(* IEC 61131-3 sources: daoli-st-library/DL_Motion (part 7) *)

(* ---- FB_DL_AxisInertiaIdent.st ---- *)
(*==============================================================================
 * 组件名称 (Component)  : FB_DL_AxisInertiaIdent
 * 所属子库 (Sublibrary) : DL_Motion
 * 当前版本 (Version)    : 1.0.0
 * 兼容性   (Platform)   : CODESYS 3.5+ / TwinCAT 3 / 汇川 InoProShop / 施耐德 Machine Expert
 *                         仅依赖 Standard.library（R_TRIG / ABS）与库内开方内核 FC_DL_SqrtEx，
 *                         零厂商私有库
 * 功能描述 (Function)   : 转动惯量与摩擦转矩在线辨识。在加速段采集 (a, T) 样本对，用最小二乘
 *                         闭式解拟合 T = J·a + Tf，得惯量 J 与摩擦转矩 Tf：
 *                         J = 〔n·ΣaT − Σa·ΣT〕/〔n·Σa² − (Σa)²〕，Tf = 〔ΣT − J·Σa〕/ n。
 *                         采样门限：|fAcc| >= fAccMin 才纳入样本；有效样本数 < nSampleMin 不出结果。
 *                         置信度：残差均方根 fRms 超 fRmsMax 时 bConfident = FALSE——**照出结果但标
 *                         不可信**（不静默丢弃，现场需要看到「拟合出来了但不可信」这个事实）。
 *                         bFreeze 为真时停止更新，fInertiaOut 保持（供调试比对）。
 * 接口     (Interface)  : 输入 fAcc 角加速度、fTorque 转矩、fAccMin 采样门限、nSampleMin 最小
 *                         样本数、fRmsMax 残差均方根上限、bEnable 使能、bFreeze 结果冻结、bReset 复位；
 *                         输出 fInertiaOut 惯量、fFrictionOut 摩擦转矩、fRms 残差均方根、
 *                         bConfident 置信标记、nSampleCount 有效样本数、eState / eCause / bError / nErrId。
 * 边界     (Boundary)   : ① 回归分母〔n·Σa² − (Σa)²〕<= DL_FLOAT_EPS 判定样本不可分（如全等
 *                         加速度），置信息级并**保持上次结果**（不清零，避免把「没算出来」错当
 *                         「惯量为 0」）；② 全部累加量用 LREAL 防精度丢失；**本件用累积量闭式解，
 *                         不使用样本环形缓冲**，故无下标越界路径（派单「环缓冲下标先判边界」
 *                         条款以零数组方式结构性满足）；
 *                         ③ 组态闸：fAccMin <= 0.0、nSampleMin = 0、fRmsMax <= 0.0 或任一浮点引脚
 *                         NaN → 故障锁存；④ 输入非有限 → 该样本剔除并计数，不污染累加量；
 *                         ⑤ R_TRIG 一枚段 0 无条件刷新（本件为纯算术拟合，无工艺相计时）；
 *                         ⑥ 故障相迁出唯一路径 = bReset 上升沿；⑦ 零全局耦合（无 GVL / 无物理地址）。
 * 解除式   (Release)    : bReset 上升沿 ∧ 组态合法 ∧ 回归分母非病态（当拍量，R240 范式）。
 *                         自证可满足（终审两式 1）：分母只依赖累加量与样本数，复位后累加量清空
 *                         即重新开始积累，加速度样本一旦分散分母即脱离病态，无恒假因子。
 * 码表     (Codes)      : 16#0004_03B7 故障级：惯量辨识故障总码（组态非法 / 输入非有限累计超限 /
 *                         非法相位），锁存至 bReset 上升沿，归因由 eCause 承载（R190 单件单总码）；
 *                         16#0004_04B7 信息级：非故障台账事件（分母病态保持上次结果 / 样本数不足）。
 *                         加码反证（R90）：二者都不改 bError、不改 eCause，且 bConfident 仍可能为真
 *                         （保持的旧结果可能高置信），若不立码则「本轮没算出新结果」不可观测，故立
 *                         一码；二者共用一码的依据是「都只要求留痕」，区分由 nSampleCount 反推。
 *                         码段说明：0004 段故障子带 03xx / 信息子带 04xx，本件取 03B7 / 04B7
 *                         （源码实扫该两槽为空，续接同子带已用最大值，未回填碎片孔洞）。
 * 开源溯源 (Origin)     : 道莅自研 clean-room（参考最小二乘闭式解与运动辨识参数域，零代码行复制；
 *                         t2-4-s7-motion 族）
 * 修订历史 (Revision)   : 2026-11-19  v1.0.0  R45 首版（批次 3 · 序号 13）
 *==============================================================================*)

TYPE E_DL_AiiState :
(
    eIdle  := 0,     // 失能或样本不足（无结果） / Idle, disabled or not enough samples
    eRun   := 10,    // 辨识运行 / Identification running
    eFault := 90     // 故障锁存相 / Fault latched phase
);
END_TYPE

TYPE E_DL_AiiCause :
(
    eNone       := 0,   // 无故障成因 / No cause
    eCfgIllegal := 1,   // 组态非法 / Illegal configuration
    eNonFinRun  := 2,   // 输入非有限累计超限 / Too many consecutive non-finite inputs
    ePhaseBad   := 3    // 非法相位兜底 / Illegal phase fallback
);
END_TYPE

FUNCTION_BLOCK FB_DL_AxisInertiaIdent
VAR_INPUT
    fAcc        : REAL := 0.0;          // 角加速度（或线加速度） [rad/s²] / Angular acceleration [rad/s2]
    fTorque     : REAL := 0.0;          // 实测转矩 [N·m] / Measured torque [N·m]
    fAccMin     : REAL := 5.0;          // 采样门限（|a| 大于该值才纳入），域 > 0.0 [rad/s²] / Sampling threshold, domain > 0.0 [rad/s2]
    nSampleMin  : UDINT := 50;          // 最小有效样本数，域 > 0 [个] / Minimum sample count, domain > 0 [pcs]
    fRmsMax     : REAL := 0.50;         // 残差均方根上限，域 > 0.0 [N·m] / Residual RMS limit, domain > 0.0 [N·m]
    bEnable     : BOOL := TRUE;         // 辨识使能 [-] / Identification enable
    bFreeze     : BOOL := FALSE;        // 结果冻结（停止更新，保持末值） [-] / Freeze results, hold last value
    bReset      : BOOL := FALSE;        // 复位命令，上升沿清故障并使累加量净重装 [-] / Reset clears fault and re-arms accumulators
END_VAR
VAR_OUTPUT
    fInertiaOut  : REAL;                // 辨识惯量（拟合斜率） [kg·m²] / Identified inertia, fitted slope [kg m2]
    fFrictionOut : REAL;                // 辨识摩擦转矩（拟合截距） [N·m] / Identified friction torque, fitted intercept [N·m]
    fRms         : REAL;                // 残差均方根（拟合优度） [N·m] / Residual RMS [N·m]
    bConfident   : BOOL;                // 置信标记（RMS 未超上限） [-] / Confident flag
    nSampleCount : UDINT;               // 当前有效样本数 [个] / Current valid sample count
    eState       : E_DL_AiiState;       // 状态出口，段 6 单点映射 / State outlet
    eCause       : E_DL_AiiCause;       // 故障成因出口（R190 归因唯一） / Fault cause outlet
    bError       : BOOL;                // 故障锁存标志 [-] / Fault latch flag
    nErrId       : UDINT;               // 事件码，0 = 无事件 / Event code, 0 = no event
END_VAR
VAR
    _eState      : E_DL_AiiState := E_DL_AiiState.eIdle;    // 内部相位（CASE 唯一写入目标） / Internal phase
    _eCause      : E_DL_AiiCause := E_DL_AiiCause.eNone;    // 故障成因锁存（锁存量） / Latched cause
    rtReset      : R_TRIG;              // 复位沿实例，段 0 无条件调用 / Reset edge
    _nSamples    : UDINT;               // 样本数（锁存量） [个] / Sample count, latched
    _fSumA       : LREAL;               // Σa（锁存量，LREAL 防精度丢失） [rad/s²] / Sum of acceleration in LREAL
    _fSumT       : LREAL;               // ΣT（锁存量） [N·m] / Sum of torque
    _fSumAA      : LREAL;               // Σa²（锁存量） [rad²/s⁴] / Sum of squared acceleration
    _fSumAT      : LREAL;               // ΣaT（锁存量） [N·m·rad/s²] / Sum of acceleration times torque
    _fSumTT      : LREAL;               // ΣT²（锁存量） [N²·m²] / Sum of squared torque
    _fDen        : LREAL;               // 回归分母 n·Σa² − (Σa)²（当拍量） [rad²/s⁴] / Regression denominator
    _fJ          : LREAL;               // 惯量拟合值（当拍量） [kg·m²] / Fitted inertia
    _fTf         : LREAL;               // 摩擦转矩拟合值（当拍量） [N·m] / Fitted friction torque
    _fSse        : LREAL;               // 残差平方和（当拍量） [N²·m²] / Residual sum of squares
    _fRmsCalc    : LREAL;               // 残差均方根计算值（当拍量） [N·m] / Computed residual RMS
    _fInertiaHold : REAL;               // 惯量保持槽（锁存量，病态时保持） [kg·m²] / Inertia hold slot, latched
    _fFricHold   : REAL;                // 摩擦保持槽（锁存量） [N·m] / Friction hold slot, latched
    _fRmsHold    : REAL;                // RMS 保持槽（锁存量） [N·m] / RMS hold slot, latched
    _bConfHold   : BOOL;                // 置信保持槽（锁存量） [-] / Confidence hold slot
    _nNonFinRun  : UDINT;               // 非有限连续计数（锁存量） [拍] / Consecutive non-finite counter
    _uSqrtErr    : UDINT;               // 开方内核错误码（当拍量） [-] / Sqrt kernel error code
    _bNonFin     : BOOL;                // 输入非有限当拍量 [-] / Non-finite input this scan
    _bCfgBad     : BOOL;                // 组态非法当拍量 [-] / Illegal configuration
    _bDenBad     : BOOL;                // 分母病态当拍量 [-] / Degenerate denominator
    _bFault      : BOOL;                // 故障锁存位（锁存量） / Latched fault bit
    _uFault      : UDINT;               // 故障码锁存（锁存量） / Latched fault code
    _uInfo       : UDINT;               // 信息码，每拍重算 / Info code, recomputed each scan
END_VAR
VAR CONSTANT
    DL_FLOAT_EPS  : LREAL := 1.0E-6;    // 浮点判零容差（分母与判据统一口径） [无量纲] / Float epsilon for zero tests
    DL_NONFIN_MAX : UDINT := 10;        // 非有限连续拍数上限 [拍] / Consecutive non-finite limit [scan]
END_VAR

(* —— 段 0：去当拍判据派生 + 沿实例无条件周期刷新 —— *)
_bNonFin := (fAcc <> fAcc) OR (fTorque <> fTorque)                                          // NaN 自反判（判等禁令唯一例外） / NaN self-reflexive tests
         OR ((fAcc - fAcc) <> (fAcc - fAcc)) OR ((fTorque - fTorque) <> (fTorque - fTorque));   // Inf 差值自减判 / Inf tests
_bCfgBad := (fAccMin <= 0.0) OR (nSampleMin = 0) OR (fRmsMax <= 0.0)                         // 组态域闸（R151 全覆盖） / Config gate
            OR (fAccMin <> fAccMin) OR (fRmsMax <> fRmsMax);                                 // 参数 NaN 判 / Parameter NaN tests
rtReset(CLK := bReset);                                                                       // 复位沿，每拍必调（R228A） / Reset edge

(* —— 段 1：单拍量预清零（锁存量不入清单，R107） —— *)
_uInfo       := 16#0000_0000;      // 信息码每拍重算 / Info recomputed every scan
nSampleCount := _nSamples;         // 样本数镜像（锁存量回放） / Sample count mirror
nErrId       := 16#0000_0000;      // 事件码缺省无事件 / Event code default none
bError       := FALSE;             // 故障标志每拍预清，故障分支同拍置位（R45 配对） / Flag preset

(* —— 段 2：复位沿（含累加量净重装）+ 组态域闸 —— *)
IF rtReset.Q THEN                                                        // 当拍复位沿 / current-scan reset edge
    _bFault := FALSE;                                                    // 清故障锁存位（锁存量） / Clear fault latch
    _uFault := 16#0000_0000;                                             // 清故障锁存码（锁存量） / Clear latched code
    _eCause := E_DL_AiiCause.eNone;                                      // 清成因（锁存量） / Clear latched cause
    _nSamples := 0;                                                      // 样本累加量净重装 / Re-arm accumulators
    _fSumA := 0.0;
    _fSumT := 0.0;
    _fSumAA := 0.0;
    _fSumAT := 0.0;
    _fSumTT := 0.0;
    _nNonFinRun := 0;                                                    // 非有限计数清空 / Clear non-finite counter
    IF _eState = E_DL_AiiState.eFault THEN
        _eState := E_DL_AiiState.eIdle;                                  // 故障相迁出唯一路径 / Sole exit from fault phase
    END_IF
END_IF
IF _bCfgBad THEN                                                         // 组态域闸 / Configuration gate
    _uFault := 16#0004_03B7;                                             // 故障级：惯量辨识故障总码 / Fault-level: identification fault code
    _bFault := TRUE;
    bError  := TRUE;                                                     // 故障标志同拍置位（R45 配对） / Error flag set same scan
    _eCause := E_DL_AiiCause.eCfgIllegal;                                // 归因：组态非法 / Cause: illegal configuration
END_IF

(* —— 段 3：样本采集（门限过滤 + 非有限剔除 + LREAL 累加） —— *)
IF (NOT _bFault) THEN
    IF _bNonFin THEN                                                     // 非有限：剔除且不污染累加量 / Non-finite sample dropped, accumulators untouched
        IF _nNonFinRun < DL_NONFIN_MAX THEN
            _nNonFinRun := _nNonFinRun + 1;
        END_IF
        _uInfo := 16#0004_04B7;                                          // 信息级：该样本剔除留痕 / Info: sample dropped
    ELSE
        _nNonFinRun := 0;                                                // 恢复有限即清连续计数 / Reset counter
        IF ABS(fAcc) >= fAccMin THEN                                     // 门限过滤（容差式） / Threshold filter
            _nSamples := _nSamples + 1;
            _fSumA  := _fSumA  + REAL_TO_LREAL(fAcc);                    // 累加 Σa / Accumulate sum of acceleration
            _fSumT  := _fSumT  + REAL_TO_LREAL(fTorque);                 // 累加 ΣT / Accumulate sum of torque
            _fSumAA := _fSumAA + REAL_TO_LREAL(fAcc) * REAL_TO_LREAL(fAcc);              // 累加 Σa² / Accumulate sum of squared acceleration
            _fSumAT := _fSumAT + REAL_TO_LREAL(fAcc) * REAL_TO_LREAL(fTorque);           // 累加 ΣaT / Accumulate cross sum
            _fSumTT := _fSumTT + REAL_TO_LREAL(fTorque) * REAL_TO_LREAL(fTorque);        // 累加 ΣT² / Accumulate sum of squared torque
        END_IF
    END_IF
END_IF
IF (NOT _bFault) AND (_nNonFinRun >= DL_NONFIN_MAX) THEN                 // 非有限累计超限置故障 / Too many non-finite inputs
    _uFault := 16#0004_03B7;
    _bFault := TRUE;
    bError  := TRUE;
    _eCause := E_DL_AiiCause.eNonFinRun;                                 // 归因：非有限累计超限 / Cause: sustained non-finite
END_IF

(* —— 段 4：最小二乘闭式解（样本够、未冻结、使能时才求解） —— *)
_bDenBad := FALSE;                                                       // 病态标记复位 / Reset degenerate marker
IF (NOT _bFault) AND bEnable AND (NOT bFreeze) AND (_nSamples >= nSampleMin) THEN
    _fDen := REAL_TO_LREAL(UDINT_TO_REAL(_nSamples)) * _fSumAA - _fSumA * _fSumA;   // 回归分母 / Regression denominator
    IF _fDen <= DL_FLOAT_EPS THEN                                        // 分母病态：样本不可分 / Degenerate denominator
        _bDenBad := TRUE;
        _uInfo := 16#0004_04B7;                                          // 信息级：分母病态，保持上次结果 / Info: degenerate, hold last result
    ELSE
        _fJ := (REAL_TO_LREAL(UDINT_TO_REAL(_nSamples)) * _fSumAT - _fSumA * _fSumT) / _fDen;   // 惯量 = 斜率 / Inertia as the slope
        _fTf := (_fSumT - _fJ * _fSumA) / REAL_TO_LREAL(UDINT_TO_REAL(_nSamples));               // 摩擦 = 截距 / Friction as the intercept
        _fSse := _fSumTT - 2.0 * _fJ * _fSumAT - 2.0 * _fTf * _fSumT
                 + _fJ * _fJ * _fSumAA + 2.0 * _fJ * _fTf * _fSumA
                 + REAL_TO_LREAL(UDINT_TO_REAL(_nSamples)) * _fTf * _fTf;                        // 残差平方和 / Residual sum of squares
        IF _fSse < 0.0 THEN                                              // 舍入误差可能给极小负值 / Rounding may make it slightly negative
            _fSse := 0.0;
        END_IF
        _fRmsCalc := FC_DL_SqrtEx(fX := _fSse / REAL_TO_LREAL(UDINT_TO_REAL(_nSamples)), eErr => _uSqrtErr);   // 委托开方内核（R140） / Delegate sqrt kernel
        _fInertiaHold := LREAL_TO_REAL(_fJ);                             // 写入保持槽（经非有限复核见段 5） / Update inertia hold slot
        _fFricHold := LREAL_TO_REAL(_fTf);                               // 写入摩擦保持槽 / Update friction hold slot
        _fRmsHold := LREAL_TO_REAL(_fRmsCalc);                           // 写入 RMS 保持槽 / Update RMS hold slot
        IF _fRmsCalc > REAL_TO_LREAL(fRmsMax) THEN
            _bConfHold := FALSE;                                         // 残差超限：标不可信但照出结果 / Mark unconfident but still publish
        ELSE
            _bConfHold := TRUE;                                          // 置信 / Confident
        END_IF
    END_IF
END_IF
IF (NOT _bFault) AND bEnable AND (NOT bFreeze) AND (_nSamples < nSampleMin) THEN
    _uInfo := 16#0004_04B7;                                              // 信息级：样本不足，不出结果 / Info: not enough samples
END_IF

(* —— 段 5：保持槽非有限复核（非有限绝不写进保持槽，R133） —— *)
IF (_fInertiaHold <> _fInertiaHold) OR (_fFricHold <> _fFricHold) OR (_fRmsHold <> _fRmsHold) THEN
    _fInertiaHold := 0.0;                                                // 非有限保持槽清零 / Zero out non-finite hold slots
    _fFricHold := 0.0;
    _fRmsHold := 0.0;
    _bConfHold := FALSE;                                                 // 置信位撤销 / Revoke confidence
END_IF

(* —— 段 6：故障解除式（R240 全当拍量） —— *)
IF rtReset.Q AND (NOT _bCfgBad) AND (NOT _bDenBad) THEN
    _bFault := FALSE;                                                    // 清故障锁存位（锁存量） / Clear fault latch
    _uFault := 16#0000_0000;                                             // 清故障锁存码（锁存量） / Clear latched code
    _eCause := E_DL_AiiCause.eNone;                                      // 清成因（锁存量） / Clear latched cause
END_IF

(* —— 段 6A：故障锁存相位迁移闸 —— *)
IF _bFault AND (_eState <> E_DL_AiiState.eFault) THEN
    _eState := E_DL_AiiState.eFault;                                     // 锁存即入故障相 / Latch enters fault phase
END_IF

(* —— 段 7：相位机（ENUM 全成员显式标签 + ELSE 兜底，R128） —— *)
CASE _eState OF

E_DL_AiiState.eIdle:
    IF (_nSamples >= nSampleMin) AND (NOT _bFault) THEN                  // 出口 1：样本够数 / Enough samples
        _eState := E_DL_AiiState.eRun;
    ELSIF _bFault THEN                                                   // 出口 2：故障锁存 / Fault latched
        _eState := E_DL_AiiState.eFault;
    END_IF

E_DL_AiiState.eRun:
    IF _nSamples < nSampleMin THEN                                       // 出口 1：样本被复位清空（前置消失，R98） / Samples re-armed
        _eState := E_DL_AiiState.eIdle;
    ELSIF _bFault THEN                                                   // 出口 2：故障锁存 / Fault latched
        _eState := E_DL_AiiState.eFault;
    END_IF

E_DL_AiiState.eFault:
    ;                                                                     // 故障相：仅段 6 复位沿可迁出 / Only the reset edge leaves this phase

ELSE
    _uFault := 16#0004_03B7;                                             // 故障级：非法相位兜底（归并总码） / Illegal-phase fallback
    _bFault := TRUE;
    bError  := TRUE;
    _eCause := E_DL_AiiCause.ePhaseBad;                                  // 归因：非法相位 / Cause: illegal phase
    _eState := E_DL_AiiState.eFault;

END_CASE

(* —— 段 8：出口单点映射（名实同源；锁存码回放；故障相安全侧） —— *)
IF _bFault THEN
    fInertiaOut  := 0.0;                                                 // 故障相惯量输出 0（不外推未知参数） / Zero inertia in fault
    fFrictionOut := 0.0;                                                 // 故障相摩擦输出 0 / Zero friction in fault
    fRms         := 0.0;                                                 // 故障相 RMS 输出 0 / Zero RMS in fault
    bConfident   := FALSE;                                               // 故障相不宣称置信 / No confidence claim in fault
ELSE
    fInertiaOut  := _fInertiaHold;                                       // 惯量出口（保持槽回放） / Inertia outlet from hold slot
    fFrictionOut := _fFricHold;                                          // 摩擦出口 / Friction outlet
    fRms         := _fRmsHold;                                           // RMS 出口 / RMS outlet
    bConfident   := _bConfHold;                                          // 置信出口 / Confidence outlet
END_IF
IF _bFault THEN
    nErrId := _uFault;                                                   // 故障锁存码回放 / Replay latched fault code
ELSE
    nErrId := _uInfo;                                                    // 信息码 / Info code
END_IF
bError := _bFault;                                                       // 故障标志与锁存同源（名实双出口，R191） / Flag from latch
eState := _eState;                                                       // 状态出口 / State outlet
eCause := _eCause;                                                       // 成因出口 / Cause outlet

END_FUNCTION_BLOCK

(* ---- FB_DL_AxisInposGuard.st ---- *)
(*
  FB_DL_AxisInposGuard  —  到位窗口判定守卫（MC_InPosition 语义 + 驻留确认） / Axis in-position guard with dwell confirm
  分类 Category : DL_Motion
  版本 Version  : 1.0.1
  来源 Source   : t1-6-plcopen — 运动守卫族零检索深化
  溯源 Origin   : clean-room 实现，MC_InPosition 语义公开借鉴，未复制任何源码行
  功能 Function : 1) 到位带双判据：|fPosition - fTarget| <= fPosBand 且 |fVelocity| <= fVelQuiet，
                  驻留 TON 持续 tDwell 后 bInpos = TRUE（tonDwell.Q 直出）；
                  2) 驻留期目标变更即复位驻留：变更判据为当拍量比较
                  ABS(fTarget - fTgtPrev) > fPosBand，禁锁存量自指；
                  3) 使能后 tWatch 内从未到位 → 故障级 03AF 锁存；
                  4) 解除式全当拍量（R240 落地），逐 BOOL 标注见段 5。
  返修记录 Rework  :
    2026-11-19  v1.0.1  R42 P0-2 中等返修：v1.0.0 监视 TON（tonWatchTo）IN 引用
                        bInpos 输出量——该量在故障相被强制 FALSE 且为本拍后段
                        计算值（跨扫描序依赖），计时基跨故障相不复位，复位后
                        残留 .Q 即刻再判 03AF（P0 派单缺陷②）。修复要点：新增
                        _bSteady 当拍量（段 0 由 _bInBand AND _bQuiet 直接承载），
                        tonWatchTo 的 IN 改为 bEnable AND (NOT _bFault) AND
                        (NOT _bSteady)——全当拍量承载，故障相与到位拍均显式
                        复位计时基；对外接口签名不变。
  边界 Boundary : ① 组态闸：fPosBand <= 0、fVelQuiet < 0、任一超时 <= 0 → 03AE 锁存；
                  ② 目标非有限或轴位置非有限 → 03B0 防御兜底锁存（NaN 自反判）；
                  ③ 驻留 TON 电平驱动：目标变更拍 IN 必断（当拍量 NOT bTgtChg 串入）；
                  ④ 无 GVL 依赖：纯引脚输入输出，无外部变量引用，无物理 IO 地址。
  依赖 Depends  : I_DL_MotionAxis（注入，不实例化）；Standard.library（TON / R_TRIG）
  码表 Error codes（Motion 段 0004，窗口 03AE~03B0 / 04AE~04B0）:
    16#0004_03AE 故障级：组态非法（到位带/静默阈/驻留/监视超时域非法），锁存至 bReset
    16#0004_03AF 故障级：驻留判据长期不满足（使能后 tWatch 未到位），锁存至 bReset
    16#0004_03B0 故障级：目标/位置非有限（防御兜底），锁存至 bReset
    16#0004_04AE 信息级：到位沿（bInpos 首次 TRUE）
    16#0004_04AF 信息级：目标变更检出（驻留复位）
    16#0004_04B0 信息级：失去到位沿（离开到位带）
  修订历史 Revision :
    2026-11-19  v1.0.0  R41 首版（批次 3 · 序号 1）
    2026-11-19  v1.0.1  R42 P0-2 中等返修（见返修记录节）
*)

FUNCTION_BLOCK FB_DL_AxisInposGuard
VAR_INPUT
    fTarget      : REAL := 0.0;       // 目标位置 [mm 或 deg]，调用方注入 / Target position injected by caller
    fPosBand     : REAL := 0.05;      // 到位带半宽 [mm 或 deg]，域 > 0 / In-position band half width
    fVelQuiet    : REAL := 1.0;       // 速度静默阈 [mm/s]，域 >= 0 / Velocity quiet threshold
    tDwell       : TIME := T#200MS;   // 驻留确认时间 [ms]，域 > 0 / Dwell confirm time
    tWatch       : TIME := T#10S;     // 未到位监视超时 [ms]，域 > 0 / Not-in-position watchdog
    bEnable      : BOOL := FALSE;     // 守卫使能 [-] / Guard enable
    bReset       : BOOL := FALSE;     // 复位，上升沿清故障锁存 / Reset edge clears fault latch
END_VAR
VAR_IN_OUT
    iAxis        : I_DL_MotionAxis;   // 运动轴引用（注入，不实例化）/ Motion axis reference
END_VAR
VAR_OUTPUT
    bInpos       : BOOL;              // 到位出口（驻留 TON 直出）[-] / In-position outlet
    bFault       : BOOL;              // 故障锁存标志 / Fault latch flag
    bError       : BOOL;              // 故障级标志（与锁存同源）/ Fault flag
    nErrId       : UDINT;             // 事件码，0 = 无事件 / Event code
END_VAR
VAR
    tonDwell     : TON;               // 驻留确认定时器，无条件周期刷新 / Dwell confirm timer
    tonWatchTo   : TON;               // 未到位监视定时器（专用超时命名），无条件刷新 / Watchdog timer
    rtReset      : R_TRIG;            // 复位沿实例，无条件刷新 / Reset edge instance
    _fTgtPrev    : REAL;              // 上拍目标快照 [mm 或 deg] / Previous target snapshot
    _bTgtChg     : BOOL;              // 目标变更当拍量 [-] / Target change current-scan flag
    _bInBand     : BOOL;              // 位置带内当拍量 [-] / In-band current-scan flag
    _bQuiet      : BOOL;              // 速度静默当拍量 [-] / Velocity-quiet current-scan flag
    _bSteady     : BOOL;              // 双判据同时成立当拍量（v1.0.1 监视 TON 计时基）/ Steady verdict current-scan flag
    _bFault      : BOOL;              // 故障锁存位（锁存量）/ Latched fault bit
    _uFault      : UDINT;             // 故障码锁存（锁存量）/ Latched fault code
    _uInfo       : UDINT;             // 信息码，每拍重算 / Transient info code
    _bInposPrev  : BOOL;              // 上拍到位镜像（到位/失位沿判据）/ Previous inpos mirror
END_VAR

(* —— 段 0：定时器与沿实例无条件周期刷新（禁置于 IF/CASE 内） —— *)
_bTgtChg := ABS(fTarget - _fTgtPrev) > fPosBand;        // 目标变更（当拍量）
_bInBand := ABS(iAxis.fPosition - fTarget) <= fPosBand; // 位置带内（当拍量）
_bQuiet := ABS(iAxis.fVelocity) <= fVelQuiet;           // 速度静默（当拍量）
_bSteady := _bInBand AND _bQuiet;                       // 双判据同立（当拍量，v1.0.1 承载监视计时基）
rtReset(CLK := bReset);                                 // 复位沿（每拍必调）
tonDwell(IN := bEnable AND _bInBand AND _bQuiet AND (NOT _bTgtChg), PT := tDwell);
                                                        // 驻留确认（目标变更拍 IN 必断，每拍必调）
tonWatchTo(IN := bEnable AND (NOT _bFault) AND (NOT _bSteady), PT := tWatch);
                                                        // 未到位监视（全当拍量承载，故障相/到位拍显式复位，v1.0.1）

(* —— 段 1：单拍量预清零（锁存量 _bFault/_uFault 不入清单，禁同拍抹除） —— *)
_uInfo := 16#0000_0000;             // 信息码每拍重算
nErrId := 16#0000_0000;             // 事件码缺省无事件

(* —— 段 2：复位沿 + 组态域闸（当拍量判据） —— *)
IF rtReset.Q THEN                   // rtReset.Q = 当拍量
    _bFault := FALSE;               // 清故障锁存位
    _uFault := 16#0000_0000;        // 清故障锁存码
END_IF
IF (fPosBand <= 0.0) OR (fVelQuiet < 0.0)
   OR (TIME_TO_DINT(tDwell) <= 0) OR (TIME_TO_DINT(tWatch) <= 0) THEN
    _uFault := 16#0004_03AE;        // 故障级：组态非法
    _bFault := TRUE;
END_IF

(* —— 段 3：非有限防御兜底（目标/位置 NaN 自反判，禁近似阈值） —— *)
IF (fTarget <> fTarget) OR (iAxis.fPosition <> iAxis.fPosition)
   OR ((fTarget - fTarget) <> (fTarget - fTarget))
   OR ((iAxis.fPosition - iAxis.fPosition) <> (iAxis.fPosition - iAxis.fPosition)) THEN
    _uFault := 16#0004_03B0;        // 故障级：非有限防御兜底
    _bFault := TRUE;
END_IF

(* —— 段 4：驻留超时锁存（判据当拍量） —— *)
IF (NOT _bFault) AND tonWatchTo.Q THEN
    _uFault := 16#0004_03AF;        // 故障级：驻留判据长期不满足
    _bFault := TRUE;
END_IF

(* —— 段 5：故障解除式（R240 落地，逐 BOOL 标注）：
     rtReset.Q = 当拍量；iAxis.bError = 当拍量；_bInBand AND _bQuiet = 当拍量。
     均不含锁存量（_bFault/_uFault），解除边真实可达。 —— *)
IF rtReset.Q AND (NOT iAxis.bError) AND _bInBand AND _bQuiet THEN
    _bFault := FALSE;               // 清故障锁存位（锁存量，仅此当拍量解除沿可清）
    _uFault := 16#0000_0000;        // 清故障锁存码（锁存量，仅本当拍量解除沿可清）
END_IF

(* —— 段 6：信息码派生（当拍量判据） —— *)
bInpos := tonDwell.Q AND (NOT _bFault);     // 到位出口（驻留 TON 直出，故障期强制 FALSE）
IF (NOT _bFault) AND bEnable THEN
    IF bInpos AND (NOT _bInposPrev) THEN
        _uInfo := 16#0004_04AE;         // 信息级：到位沿
    END_IF
    IF _bTgtChg AND bInpos THEN
        _uInfo := 16#0004_04AF;         // 信息级：目标变更检出（驻留已复位）
    END_IF
    IF (NOT bInpos) AND _bInposPrev THEN
        _uInfo := 16#0004_04B0;         // 信息级：失去到位沿
    END_IF
END_IF

(* —— 段 7：出口单点映射（锁存码回放，禁同拍抹除） —— *)
IF _bFault THEN
    nErrId := _uFault;              // 故障锁存码回放
    bInpos := FALSE;                // 故障期到位强制 FALSE（安全侧）
ELSE
    nErrId := _uInfo;               // 信息码
END_IF
bFault := _bFault;                  // 锁存位出口
bError := _bFault;                  // 故障标志与锁存位同源
_bInposPrev := bInpos;              // 到位沿判据快照
_fTgtPrev := fTarget;               // 上拍目标快照（段末统一写）

END_FUNCTION_BLOCK

(* ---- FB_DL_AxisJerkLimitCheck.st ---- *)
(*
  Name        : FB_DL_AxisJerkLimitCheck
  Category    : DL_Motion
  Version     : 1.0.0
  Purpose     : 加加速度（jerk）指令合法性检查与钳位：由速度指令序列二次差分得加速度与 jerk，jerk 越限时把本拍速度指令回退到「上一拍加速度 ± jerk 上限」允许的取值，防高速贴装冲击；/ Check and clamp jerk of a velocity command sequence: derive acceleration and jerk by successive differences, and when jerk exceeds the limit back off the velocity command to the value permitted by the jerk-limited acceleration
  溯源        : 借 t1-6-plcopen·limits 的分类/参数域组织，clean-room 实现
  Boundary    : ① 组态闸：扫描周期 <= T#0S / jerk 上限 <= eps / 加速度上限 <= eps / 速度上限 <= eps → 锁存故障；
                ② 二次差分除子 dt 秒值在组态闸后使用，且使用前再判 > eps（双保险）；
                ③ 非有限速度指令该拍直通不钳位（保持上拍状态量，不作伪钳位）；
                ④ 输出速度钳到 [-fVelMax, +fVelMax]（双侧直比，不用 ABS 单侧）；
                ⑤ 本件只改「指令」，不参与位置环闭环；钳位生效即置 bLimited，供上层记录。
*)
TYPE E_DL_AjcState :
(
    eIdle  := 0,                             (* 未使能 / Disabled *)
    eChk   := 10,                            (* 检查运行 / Checking *)
    eFault := 90                             (* 故障锁存相 / Fault latched *)
);
END_TYPE

TYPE E_DL_AjcCause :
(
    eNone       := 0,                        (* 无故障成因 / No cause *)
    eCfgIllegal := 1,                        (* 组态非法：周期/限值越域 / Illegal config *)
    ePhaseBad   := 2                         (* 非法相位兜底 / Illegal phase fallback *)
);
END_TYPE

FUNCTION_BLOCK FB_DL_AxisJerkLimitCheck
VAR_INPUT
    fVelCmd   : REAL := 0.0;                 (* 原始速度指令 [mm/s] / Raw velocity command *)
    tScan     : TIME := T#4MS;               (* 指令更新周期，域 > T#0S [ms] / Command update period, > 0 *)
    fJerkMax  : REAL := 1.0E5;               (* 允许 jerk 上限，域 > 0 [mm/s³] / Allowed jerk limit, > 0 *)
    fAccMax   : REAL := 1.0E4;               (* 允许加速度上限，域 > 0 [mm/s²] / Allowed acceleration limit, > 0 *)
    fVelMax   : REAL := 2000.0;              (* 速度双向限幅，域 > 0 [mm/s] / Symmetric velocity limit, > 0 *)
    bEnable   : BOOL := TRUE;                (* 检查使能 [-] / Enable *)
    bReset    : BOOL := FALSE;               (* 复位命令，上升沿清状态量与标志 [-] / Reset command *)
END_VAR
VAR_OUTPUT
    fVelOut   : REAL;                        (* 钳位后速度指令 [mm/s] / Clamped velocity command *)
    fAcc      : REAL;                        (* 本拍实测加速度 [mm/s²] / Measured acceleration this scan *)
    fJerk     : REAL;                        (* 本拍实测 jerk [mm/s³] / Measured jerk this scan *)
    bLimited  : BOOL;                        (* 本拍钳位生效 [-] / Clamp applied this scan *)
    bVelClamp : BOOL;                        (* 本拍速度限幅生效（与 jerk 钳位分开归因）[-] / Velocity clamp applied *)
    eState    : E_DL_AjcState;               (* 状态出口 / State outlet *)
    eCause    : E_DL_AjcCause;               (* 故障成因出口（R190 归因唯一） / Fault cause outlet *)
    bError    : BOOL;                        (* 故障锁存标志 [-] / Fault latch flag *)
END_VAR
VAR
    _eState  : E_DL_AjcState := E_DL_AjcState.eIdle;     (* 内部相位（CASE 唯一写入目标） / Internal phase *)
    _eCause  : E_DL_AjcCause := E_DL_AjcCause.eNone;     (* 故障成因锁存量 / Latched cause *)
    rtReset  : R_TRIG;                       (* 复位沿实例，段 0 无条件调用 / Reset edge instance *)
    _bFault  : BOOL;                         (* 故障锁存位 / Latched fault bit *)
    _bCfgBad : BOOL;                         (* 组态非法当拍量 / Illegal config this scan *)
    _bFinite : BOOL;                         (* 输入有限性当拍量 / Input finiteness *)
    _fDtSec  : REAL;                         (* 周期秒值，域 > eps [s] / Period in seconds *)
    _fVelPrev: REAL;                         (* 上拍（钳位后）速度快照 [mm/s] / Previous clamped velocity *)
    _fAccPrev: REAL;                         (* 上拍加速度快照 [mm/s²] / Previous acceleration *)
    _fAccNew : REAL;                         (* 本拍加速度（由速度差分）[mm/s²] / New acceleration *)
    _fJerkNew: REAL;                         (* 本拍 jerk（由加速度差分）[mm/s³] / New jerk *)
    _fAccLim : REAL;                         (* jerk 受限后允许的加速度 [mm/s²] / Jerk-limited acceleration *)
    _fVelTgt : REAL;                         (* 未限幅的目标速度 [mm/s] / Target velocity before clamp *)
    _fVelCl  : REAL;                         (* 限幅后速度中间量 [mm/s] / Clamped velocity intermediate *)
END_VAR
VAR CONSTANT
    DL_AJC_EPS : REAL := 1.0E-6;             (* 判零容差（REAL 量级，含 dt/限值）[-] / Epsilon *)
END_VAR

(* —— 段 0：当拍判据派生 + 实例无条件刷新（R228A） —— *)
_fDtSec := TIME_TO_LREAL(tScan) / 1000.0;                                      (* 周期秒化（除子常量 1000） / Period to seconds *)
_bCfgBad := NOT (tScan > T#0S)                                                 (* 周期正域闸（二次差分除零前置） / Period gate *)
            OR (fJerkMax <= DL_AJC_EPS)                                        (* jerk 上限正域闸 / Jerk gate *)
            OR (fAccMax <= DL_AJC_EPS)                                         (* 加速度上限正域闸 / Acc gate *)
            OR (fVelMax <= DL_AJC_EPS);                                        (* 速度上限正域闸 / Velocity gate *)
rtReset(CLK := bReset);                                                        (* 复位沿每拍必调 / Reset edge every scan *)
_bFinite := (fVelCmd = fVelCmd) AND ((fVelCmd - fVelCmd) = (fVelCmd - fVelCmd));   (* NaN 自反 + Inf 差判联合闸 / NaN and Inf gate *)

(* —— 段 1：单拍量预清零（R107） —— *)
bLimited := FALSE;                                                             (* jerk 钳位预清 / Jerk clamp preset *)
bVelClamp := FALSE;                                                            (* 速度限幅预清 / Velocity clamp preset *)
fVelOut := fVelCmd;                                                            (* 出口缺省直通（未命中钳位分支时语义） / Outlet default passthrough *)

(* —— 段 2：复位沿处理（作用域：清故障 + 清差分状态量 + 迁 eIdle，R283 逐项声明） —— *)
IF rtReset.Q THEN
    _bFault := FALSE;                                                          (* 清故障锁存 / Clear fault *)
    _eCause := E_DL_AjcCause.eNone;                                            (* 清成因 / Clear cause *)
    _fVelPrev := 0.0;                                                          (* 清速度快照（复位后从静止起算） / Clear velocity snapshot *)
    _fAccPrev := 0.0;                                                          (* 清加速度快照 / Clear acceleration snapshot *)
    fVelOut := 0.0;                                                            (* 出口归零（静止态） / Outlet zeroed *)
    fAcc := 0.0;                                                               (* 清加速度出口 / Clear acc outlet *)
    fJerk := 0.0;                                                              (* 清 jerk 出口 / Clear jerk outlet *)
    _eState := E_DL_AjcState.eIdle;                                            (* 迁未使能相 / Back to idle *)
END_IF

(* —— 段 3：组态故障锁存（锁存至复位沿，R189） —— *)
IF _bCfgBad AND NOT _bFault THEN
    _bFault := TRUE;                                                           (* 锁存故障位 / Latch fault *)
    _eCause := E_DL_AjcCause.eCfgIllegal;                                      (* 成因：组态非法 / Cause: illegal config *)
    _eState := E_DL_AjcState.eFault;                                           (* 同步迁故障相 / Migrate to fault *)
END_IF

(* —— 段 4：CASE 主状态机（ELSE 兜底迁 eFault，红线 6） —— *)
CASE _eState OF
    E_DL_AjcState.eIdle:                                                       (* 未使能：指令直通，不检查 / Disabled *)
        fVelOut := fVelCmd;                                                    (* 直通（不出钳位） / Passthrough *)
        _fVelPrev := fVelCmd;                                                  (* 快照跟随，避免重使能首拍虚假 jerk / Track snapshot *)
        _fAccPrev := 0.0;                                                      (* 加速度快照清零 / Acc snapshot cleared *)
        IF bEnable AND NOT _bFault THEN
            _eState := E_DL_AjcState.eChk;                                     (* 使能进入检查 / Enter checking *)
        END_IF
    E_DL_AjcState.eChk:                                                        (* 检查相：差分求 acc/jerk + 越限钳位 / Checking *)
        IF NOT bEnable THEN
            _eState := E_DL_AjcState.eIdle;                                    (* 失能回未使能 / Back to idle *)
        ELSIF _bFinite AND (_fDtSec > DL_AJC_EPS) THEN
            _fAccNew := (fVelCmd - _fVelPrev) / _fDtSec;                       (* 加速度 = Δv/dt（除子已过闸）[mm/s²] / Acceleration, divisor gated *)
            _fJerkNew := (_fAccNew - _fAccPrev) / _fDtSec;                     (* jerk = Δa/dt（除子已过闸）[mm/s³] / Jerk, divisor gated *)
            fAcc := _fAccNew;                                                  (* 加速度出口 / Acc outlet *)
            fJerk := _fJerkNew;                                                (* jerk 出口 / Jerk outlet *)
            IF _fJerkNew > fJerkMax THEN
                _fAccLim := _fAccPrev + fJerkMax * _fDtSec;                    (* 正向越限：加速度只许升到上限步长 / Positive: limit acc rise *)
                bLimited := TRUE;                                              (* 钳位生效 / Clamp applied *)
            ELSIF _fJerkNew < (-fJerkMax) THEN
                _fAccLim := _fAccPrev - fJerkMax * _fDtSec;                    (* 负向越限：加速度只许降到下限步长 / Negative: limit acc fall *)
                bLimited := TRUE;                                              (* 钳位生效 / Clamp applied *)
            ELSE
                _fAccLim := _fAccNew;                                          (* 未越限：沿用实测加速度 / No clamp *)
            END_IF
            IF _fAccLim > fAccMax THEN
                _fAccLim := fAccMax;                                           (* 加速度上限双侧直比 / Acc upper clamp *)
                bLimited := TRUE;                                              (* 计入钳位归因 / Count as clamp *)
            ELSIF _fAccLim < (-fAccMax) THEN
                _fAccLim := -fAccMax;                                          (* 加速度下限双侧直比 / Acc lower clamp *)
                bLimited := TRUE;                                              (* 计入钳位归因 / Count as clamp *)
            END_IF
            _fVelTgt := _fVelPrev + _fAccLim * _fDtSec;                        (* 由受限加速度重建本拍速度指令 / Rebuild velocity from limited acc *)
            _fVelCl := _fVelTgt;                                               (* 限幅前中间量 / Intermediate before clamp *)
            IF _fVelCl > fVelMax THEN
                _fVelCl := fVelMax;                                            (* 速度上限钳位（双侧直比，禁 ABS 单侧） / Velocity upper clamp *)
                bVelClamp := TRUE;                                             (* 限幅归因独立（R190） / Velocity clamp cause *)
            ELSIF _fVelCl < (-fVelMax) THEN
                _fVelCl := -fVelMax;                                           (* 速度下限钳位 / Velocity lower clamp *)
                bVelClamp := TRUE;                                             (* 限幅归因独立 / Velocity clamp cause *)
            END_IF
            fVelOut := _fVelCl;                                                (* 钳位后指令出口 / Clamped command outlet *)
            _fVelPrev := _fVelCl;                                              (* 快照推进为钳位后值（下拍差分基准） / Advance snapshot *)
            _fAccPrev := _fAccLim;                                             (* 加速度快照推进为受限值 / Advance acc snapshot *)
        END_IF                                                                 (* 非有限/周期退化：直通不钳位（边界③） / Passthrough *)
    E_DL_AjcState.eFault:                                                      (* 故障相：冻结保持末值，仅复位沿出 / Fault *)
        ;                                                                      (* 锁存回放（R28） / Replay from latch *)
    ELSE                                                                       (* 非法相位兜底迁安全态 / Illegal phase fallback *)
        _eState := E_DL_AjcState.eFault;                                       (* 迁故障相 / To fault *)
        _bFault := TRUE;                                                       (* 同步锁存 / Latch *)
        _eCause := E_DL_AjcCause.ePhaseBad;                                    (* 成因：非法相位 / Cause: illegal phase *)
END_CASE

(* —— 段 5：出口映射（bError/eState 同源，R191） —— *)
bError := _bFault;                                                             (* 故障标志镜像 / Fault flag mirror *)
eState := _eState;                                                             (* 状态出口 / State outlet *)
eCause := _eCause;                                                             (* 成因出口 / Cause outlet *)
END_FUNCTION_BLOCK

(* ---- FB_DL_AxisJogController.st ---- *)
(*==============================================================================
 * 组件名称 (Component)  : FB_DL_AxisJogController
 * 所属子库 (Sublibrary) : DL_Motion
 * 当前版本 (Version)    : 1.0.0
 * 组件分类 (Category)   : 功能块（FUNCTION_BLOCK）· 轴点动操作器 · 工艺上层件
 * 兼容性   (Platform)   : CODESYS 3.5 / TwinCAT 3 / 汇川 InoProShop / Schneider
 *                         Machine Expert；仅依赖 Standard.library（TON / R_TRIG /
 *                         MIN / MAX / ABS），零厂商方言
 * 功能描述 (Function)   : 单轴点动操作器，经 I_DL_MotionAxis 接口引用驱动
 *                         轴体（依赖注入，不关心实现块品牌）。点动语义：
 *                         长按低速、按住高速选择且延时到自动升高速、松开
 *                         即受控停止；升/降速均走轴接口速度域限幅斜坡，
 *                         不做阶跃。软限位拦截独立于轴组态，便于现场收紧：
 *                         进入制动距离警戒区强制降为低速，限位处拒绝继续。
 * 设计要点 (Key notes)  : ① 双向同按 → 停止 + 信息级 0004_0102（安全侧
 *                           「不猜」，两方向都不执行）；
 *                         ② iAxis 不在 eStandstill/eContinuousMotion → 点动
 *                           指令拒绝（含 eStopping/eErrorStop 门禁）；
 *                         ③ 制动距离 fBrakeDist = fVel²/(2·fAcc) 现算（S-2
 *                           软限位预判语义的简化版），fAcc 有参数下限兜底
 *                           防除零；
 *                         ④ 参数对调自修复（公约 0.6）：fJogSlow > fJogFast
 *                           对调、限位对倒置对调，信息级 0004_0103。
 * 规格偏离留档 (R11)    : 规格引脚表未列 uErrorId，但信息级出码（0102/0103/
 *                         0105）必须有可观察出口，故补充 uErrorId : UDINT
 *                         输出引脚（信息级专用，无故障锁存语义）。
 * 开源溯源 (Origin)     : s7-motion。仅提取 S7-1500 Motion Control 手册公开
 *                         的点动工艺语义（低速/高速点动、延时切换）与接口
 *                         参数域；实现与命名 100% 自有 clean-room。
 * 验收向量 (Acceptance) :
 *   V1 正常链：bJogPos 按住 → iAxis 进入 eContinuousMotion 正向低速；
 *      bFastSelect 按住且 tFastDelay 到 → 升高速；松开 → iAxis.Stop()；
 *   V2 双向同按：bJogPos+bJogNeg → 停止请求 + 信息级 0004_0102；
 *   V3 软限位拦截：正向点动接近 fSoftLimitPos 制动距离内 → 强制低速；
 *      到限位 → 停止请求 + 信息级 0004_0105；
 *   V4 参数对调：fJogSlow=50 / fJogFast=5 → 对调生效 + 信息级 0004_0103；
 *   V5 状态门禁：iAxis.eState = eErrorStop → 点动指令被拒，轴状态不变。
 * 故障码表 (Error codes):
 *   16#0004_0102【信息级】双向点动冲突 / 16#0004_0103【信息级】参数对调
 *   或兜底修复 / 16#0004_0105【信息级】软限位预判停车（与 FB_DL_SingleAxis
 *   同码同义，点动与连续运动共用）。
 * 修订历史 (Revision)   :
 *   2026-11-15  v1.0.0  首版入库（Round 05 · DL_Motion 开库）
 *============================================================================*)

(*-----------------------------------------------------------------------------
 * 调用示例 (Instance guide)：
 *   fbJog.iAxis := fbAxis;                        // 接口依赖注入（注入实现块实例）
 *   fbJog(bJogPos := bBtnUp, bJogNeg := bBtnDown, // 周期调用
 *         bFastSelect := bBtnFast, fJogSlow := 5.0, fJogFast := 50.0);
 *   手轮/按键电平直接接 bJogPos/bJogNeg；松开即停，无需上层编排停止时序。
 *   点动软限位独立于轴组态：现场试机时可临时收紧 fSoftLimitPos/Neg。
 *----------------------------------------------------------------------------*)

(*-----------------------------------------------------------------------------
 * 常见误用与现场提示 (Field notes)：
 *   1 点动速度变化走轴的速度域斜坡（MoveVelocity 改速语义），但加减速
 *     由 fAcc 单参数承担，现场要求的"点动要跟手"请把 fAcc 适当调大，
 *     不要去改轴的组态参数。
 *   2 高速切换是"按住 bFastSelect 且已按方向键满 tFastDelay"，不是按
 *     高速键的边沿；想瞬切高速的工位把 tFastDelay 设为 T#0MS 即可
 *     （TON 零延时当拍满足）。
 *   3 本块不做任何传感器/安全件防抖，急停与安全门请走 bProcessAbort /
 *     驱动层安全链，不要指望点动块拦截。
 *   4 点动软限位与轴组态软限位是两道独立防线，两者取交集生效；现场
 *     收紧本块限位不会影响程序自动运行的轴组态限位。
 *----------------------------------------------------------------------------*)
FUNCTION_BLOCK FB_DL_AxisJogController
VAR_INPUT
    bJogPos        : BOOL := FALSE;      // 正向点动（Jog forward），电平生效
    bJogNeg        : BOOL := FALSE;      // 负向点动（Jog backward），电平生效
    fJogSlow       : REAL := 5.0;        // 低速点动速度（Slow jog velocity）[mm/s]
    fJogFast       : REAL := 50.0;       // 高速点动速度（Fast jog velocity）[mm/s]
    bFastSelect    : BOOL := FALSE;      // 高速选择（Fast select），TRUE 且按住 ≥ tFastDelay 自动切高速
    tFastDelay     : TIME := T#1S;       // 低→高速切换延时（Fast switch delay）
    fSoftLimitPos  : REAL := 1000000.0;  // 点动软限位上限（Jog soft limit high）[mm]，独立于轴组态
    fSoftLimitNeg  : REAL := -1000000.0; // 点动软限位下限（Jog soft limit low）[mm]
    fAcc           : REAL := 1000.0;     // 点动加减速度（Jog acceleration）[mm/s²]
END_VAR
VAR_IN_OUT
    iAxis          : I_DL_MotionAxis;    // 轴接口引用（Axis reference），由上层注入实现块实例
END_VAR
VAR_OUTPUT
    uErrorId       : UDINT := 0;         // 末次信息级事件码（Last info code），规格外补充引脚（见头注 R11 留档）
END_VAR
VAR
    bJogging       : BOOL := FALSE;      // 点动进行中（Jog active）
    bStopReq       : BOOL := FALSE;      // 内部停止请求（Internal stop request）
    bAxisOk        : BOOL := FALSE;      // 轴状态可用标志（Axis state usable），eStandstill/eContinuousMotion 为 TRUE
    iJogMode       : INT := 0;           // 点动模式裁决值（Jog mode decision）：0 停止/1 正向/2 负向/3 冲突
    fVelSel        : REAL := 5.0;        // 生效点动速度（Selected jog speed）[mm/s]
    fVelCmd        : REAL := 0.0;        // 本拍点动速度指令（Jog velocity command）[mm/s]，带符号
    fSlow          : REAL := 5.0;        // 生效低速（Effective slow speed）[mm/s]，对调修复后
    fFast          : REAL := 50.0;       // 生效高速（Effective fast speed）[mm/s]，对调修复后
    fAccEff        : REAL := 1000.0;     // 生效加减速度（Effective acceleration）[mm/s²]
    fLimPos        : REAL := 1000000.0;  // 生效点动软限位上限（Effective jog limit high）[mm]
    fLimNeg        : REAL := -1000000.0; // 生效点动软限位下限（Effective jog limit low）[mm]
    fBrakeDist     : REAL := 0.0;        // 制动距离（Braking distance）[mm]
    fDistToLim     : REAL := 0.0;        // 沿点动方向距限位距离（Distance to limit）[mm]
    tonFast        : TON;                // 低→高速切换延时定时器（Fast switch delay timer）
    rtrigStop      : R_TRIG;             // 停止请求沿检测（Rising edge of stop request）
END_VAR
VAR CONSTANT
    DL_JOG_INF_MAX  : REAL := 1.0E30;    // 有限值判定幅值上限（Finite-value magnitude bound）[mm]
    DL_JOG_EPS      : REAL := 1.0E-6;    // 浮点判零容差（Float zero tolerance）[mm]
    DL_JOG_ACC_FLOOR : REAL := 1.0E-3;   // 加速度参数下限兜底（Acceleration parameter floor）[mm/s²]
END_VAR

METHOD DispatchJog : BOOL
VAR_INPUT
    bPositive : BOOL;                    // 点动方向（Jog direction），TRUE=正向
END_VAR
DispatchJog := FALSE;
// 速度选择：长按低速，按住高速选择且延时到自动升高速
fVelSel := fSlow;
IF bFastSelect AND tonFast.Q THEN
    fVelSel := fFast;
END_IF
// 软限位预判：制动距离内强制低速，限位处拒绝继续
IF bPositive THEN
    fDistToLim := fLimPos - iAxis.fPosition;          // 正向距限位 [mm]
ELSE
    fDistToLim := iAxis.fPosition - fLimNeg;          // 负向距限位 [mm]
END_IF
fBrakeDist := (fVelSel * fVelSel) / (2.0 * fAccEff);  // 制动距离 [mm]，fAccEff 有下限防除零
IF fDistToLim <= DL_JOG_EPS THEN
    bStopReq := TRUE;                    // 已在限位：拒绝继续点动
    uErrorId := 16#0004_0105;
    RETURN;
ELSIF fDistToLim <= fBrakeDist THEN
    fVelSel := fSlow;                    // 警戒区内强制降为低速（预判语义简化版）
END_IF
// 发速度指令：带符号速度走轴接口速度域限幅斜坡，不做阶跃
IF bPositive THEN
    fVelCmd := fVelSel;
ELSE
    fVelCmd := -fVelSel;
END_IF
IF iAxis.MoveVelocity(fVelCmd, fAccEff) THEN
    bJogging := TRUE;
    DispatchJog := TRUE;
END_IF
    END_METHOD

// 段 1｜定时器/沿检测无条件周期刷新（R7 红线，严禁置于分支内）
tonFast(CLK := (bJogPos XOR bJogNeg) AND bFastSelect AND (NOT bStopReq), PT := tFastDelay);
rtrigStop(CLK := bStopReq);

// 段 2｜接口引用有效性防御：未注入轴引用则直接退出（不产生误动作）
IF iAxis = 0 THEN
    bJogging := FALSE;
    RETURN;
END_IF

// 段 3｜轴状态门禁：仅待机/连续运动两态可点动（eStopping/eErrorStop 拒绝）
bAxisOk := (iAxis.eState = E_DL_AxisState.eStandstill) OR (iAxis.eState = E_DL_AxisState.eContinuousMotion);

// 段 4｜参数防御与对调自修复（公约 0.6/0.8）：信息级码，不锁存
IF (fJogSlow <> fJogSlow) OR (fJogFast <> fJogFast) OR (fJogSlow <= DL_JOG_EPS) OR (fJogFast <= DL_JOG_EPS)
   OR (fJogSlow > DL_JOG_INF_MAX) OR (fJogFast > DL_JOG_INF_MAX) THEN
    fSlow := 5.0;                        // 非有限/非法低速兜底 [mm/s]
    fFast := 50.0;                       // 非有限/非法高速兜底 [mm/s]
    uErrorId := 16#0004_0103;
ELSIF fJogSlow > fJogFast THEN
    fSlow := fJogFast;                   // 低/高速对调修复（Swap repair）
    fFast := fJogSlow;
    uErrorId := 16#0004_0103;
ELSE
    fSlow := fJogSlow;
    fFast := fJogFast;
END_IF
IF (fAcc <> fAcc) OR (fAcc <= DL_JOG_ACC_FLOOR) OR (fAcc > DL_JOG_INF_MAX) THEN
    fAccEff := 1000.0;                   // 非法加速度兜底 [mm/s²]，防除零
    uErrorId := 16#0004_0103;
ELSE
    fAccEff := fAcc;
END_IF
IF fSoftLimitPos < fSoftLimitNeg THEN
    fLimPos := fSoftLimitNeg;            // 点动限位对倒置对调修复（Swap repair）
    fLimNeg := fSoftLimitPos;
    uErrorId := 16#0004_0103;
ELSE
    fLimPos := fSoftLimitPos;
    fLimNeg := fSoftLimitNeg;
END_IF

// 段 5｜点动模式裁决：双向冲突/松开/正常三分支（安全侧不猜）
IF bJogPos AND bJogNeg THEN
    iJogMode := 3;                       // 双向同按：冲突模式
ELSIF (NOT bJogPos) AND (NOT bJogNeg) THEN
    iJogMode := 0;                       // 松开：停止模式
ELSIF bAxisOk THEN
    IF bJogPos THEN iJogMode := 1; ELSE iJogMode := 2; END_IF   // 正向/负向点动
ELSE
    iJogMode := 0;                       // 轴态不可用：按松开处理
END_IF

// 段 6｜点动决策机（CASE+ELSE 兜底）
CASE iJogMode OF
    0:                                   // 停止模式：等待停止沿
        bJogging := FALSE;
    1:                                   // 正向点动
        IF NOT DispatchJog(bPositive := TRUE) THEN
            bStopReq := TRUE;            // 轴拒绝受理 → 转停止
        END_IF
    2:                                   // 负向点动
        IF NOT DispatchJog(bPositive := FALSE) THEN
            bStopReq := TRUE;
        END_IF
    3:                                   // 冲突模式：两方向都不执行
        bStopReq := TRUE;
        uErrorId := 16#0004_0102;
        bJogging := FALSE;
ELSE
    // 非法模式兜底
    iJogMode := 0;
END_CASE

// 段 7｜停止沿执行：松开/冲突/限位停车 → 调用轴受控停止（MC_Stop 语义），
//      消费后才清标志，保证 R_TRIG 能捕获到电平（沿在本拍段 1 已建立）
IF rtrigStop.Q THEN
    iAxis.Stop();
    bStopReq := FALSE;
END_IF

(*-----------------------------------------------------------------------------
 * 方法实现（METHOD）：点动派发子过程，速度选择 + 软限位预判 + 发速度指令
 * 三步串行，供主体点动决策机调用，正/负向共用一套逻辑。
 *-----------------------------------------------------------------------------*)

END_FUNCTION_BLOCK

(* ---- FB_DL_AxisLimitRecovery.st ---- *)
(*
  FB_DL_AxisLimitRecovery  —  硬限位触发后的脱离恢复顺控 / Hard-limit trigger back-off recovery sequence
  分类 Category : DL_Motion
  码位 Code     : 16#04_0_A7
  段位说明      : A6 格由 FB_DL_CamOverrideTrim 启用，本件启用相邻 A7 格（一件一码）
  版本 Version  : 1.0.1
  来源 Source   : t1-6-plcopen — 硬限位恢复顺控待挖项落地
  溯源 Origin   : clean-room 实现，PLCopen 恢复语义公开借鉴，未复制任何源码行
  功能 Function : 1) 七相顺控 Idle→Judge→Backoff→Confirm→Reenable→Done，判限位方向 → 低速反向
                  脱离 → 脱离确认 → 重新使能放行；
                  2) 判向：bLimPos 触发反向退、bLimNeg 触发正向退、双限同拍判组态/硬件故障；
                  3) 脱离确认双判据：限位开关释放 AND FB_DL_AxisInPosMonitor 稳定到位（防半脱假通过）；
                  4) 放行再使能：CmdReset → Enable(TRUE)，等 bEnabled 落定才进 Done。
  边界 Boundary : ① 与 FB_DL_SoftLimitGuard（软限位制动预判）分工：那件管预防，本件管硬限位已触发后的恢复；
                  与 FB_DL_TorqueLimitControl（达限即限）分工：那件管力矩限制本身；
                  ② 脱离移动经 I_DL_MotionAxis.MoveRelative 单发下发（进入相拍一次，方法内受理去重）；
                  ③ R228-A 达标声明：四只超时 TON 均单相独占（IN 为单相等式），跨相迁移拍 IN 必断；
                  ④ R228-B 达标声明（R41 P0-1 返修后逐字自证，与段 4 实现逐字对照）：
                  eFault 迁出 = rtReset.Q（当拍量） AND NOT iAxis.bError（当拍量）
                  AND NOT (bLimPos AND bLimNeg)（当拍量）——三个子条件全部为当拍量，
                  零锁存量自指（R240 修复点）；可满足性：双限不同拍触发（正常工况）
                  AND 轴无报警 AND 复位沿到达，迁出边真实可达，无恒假子式；
                  ⑤ 起始时无限位触发：置信息级码并停留 Idle（不做无意义移动）。
  依赖 Depends  : I_DL_MotionAxis（注入，不实例化）；FB_DL_AxisInPosMonitor（实例化，引脚按 registry 实名）
  码表 Error codes（本件格 04_0_A7，子码步进 +0x100）:
    16#0004_01A7 信息级：恢复完成（Done 相）
    16#0004_02A7 故障级：双限位同拍触发（组态/硬件矛盾），锁存至复位
    16#0004_03A7 故障级：段超时（Judge/Backoff/Confirm/Reenable 各相独立计时），锁存至复位
    16#0004_04A7 故障级：轴故障锁存（iAxis.bError），锁存至复位
    16#0004_05A7 故障级：状态机落 ELSE 兜底（非法相位 ID），锁存至复位
    16#0004_06A7 信息级：起始时无限位触发（无需恢复，停留 Idle）
    16#0004_07A7 故障级：组态非法（距离/速度/加速度/容差/超时域非法），锁存至复位

  修订历史 Revision :
    2026-11-19  v1.0.0  R39 首版（批次 2 · 序号 8）
    2026-11-19  v1.0.1  R40 5 抽终审挂账（不改逻辑）：⚠ 段 4 解除式「rtReset.Q AND NOT _bFault」
                  引用锁存位自身，锁存后恒假 → eFault 永久锁死（R28-1 典型反例）；修复方向 = 改按
                  当前条件判定（NOT iAxis.bError AND NOT (bLimPos AND bLimNeg)），返修轮处理。
    2026-11-19  v1.0.1  R41 P0-1 返修实施：段 4 解除式重构为「rtReset.Q AND NOT iAxis.bError
                  AND NOT (bLimPos AND bLimNeg)」，全部当拍量、零锁存量自指；每个解除式 BOOL
                  已在段 4 逐个标注锁存量/当拍量；头注释④自证句与实现逐字对照。
*)

TYPE E_DL_AxlRecState :
(
    eIdle     := 0,    // 空闲：等恢复指令 / Idle, waiting for recovery command
    eJudge    := 10,   // 判向：确定脱离方向 / Judge, determine back-off direction
    eBackoff  := 20,   // 脱离：低速反向移动 / Backoff, low-speed reverse move
    eConfirm  := 30,   // 确认：限位释放 + 稳定到位 / Confirm, limit released and settled
    eReenable := 40,   // 放行：复位报警 + 再使能 / Reenable, reset alarm and power on
    eDone     := 50,   // 完成：恢复落定 / Done
    eFault    := 90    // 故障：双限/超时/轴故障锁定 / Fault, latched
);
END_TYPE

FUNCTION_BLOCK FB_DL_AxisLimitRecovery
VAR_INPUT
    bStartRec    : BOOL := FALSE;     // 恢复指令（上升沿）/ Recovery start command
    bLimPos      : BOOL := FALSE;     // 正向硬限位开关，TRUE = 已触发 [-] / Positive hard limit switch, TRUE = tripped
    bLimNeg      : BOOL := FALSE;     // 负向硬限位开关，TRUE = 已触发 [-] / Negative hard limit switch, TRUE = tripped
    fBackoffDist : REAL := 5.0;       // 脱离距离 [mm]，域 (0, 10000] / Back-off distance
    fBackoffVel  : REAL := 2.0;       // 脱离速度 [mm/s]，域 (0, 1000] / Back-off velocity
    fBackoffAcc  : REAL := 50.0;      // 脱离加/减速度 [mm/s²]，域 > 0 / Back-off acceleration
    fPosTol      : REAL := 0.05;      // 确认相位置窗半宽 [mm]，域 > 0 / Confirm-phase position tolerance
    fVelTol      : REAL := 1.0;       // 确认相速度阈 [mm/s]，域 > 0 / Confirm-phase velocity threshold
    tPhaseTo     : TIME := T#10S;     // 单相超时 [ms]，域 > 0 / Per-phase timeout
    bReset       : BOOL := FALSE;     // 复位（eFault 迁出沿之一）/ Reset, fault exit edge
END_VAR
VAR_OUTPUT
    eState       : E_DL_AxlRecState;  // 状态出口，段尾单点映射 / State outlet
    bRecovered   : BOOL;              // 恢复完成锁存（Done 相置位，Idle 相清除）/ Recovered latch
    bBackDirNeg  : BOOL;              // 本次脱离方向（TRUE = 负向）/ Back-off direction of this recovery
    nErrId       : UDINT;             // 事件码，0 = 无事件 / Event code
END_VAR
VAR_IN_OUT
    iAxis : I_DL_MotionAxis;          // 运动轴引用（注入，不实例化）/ Motion axis reference
END_VAR
VAR
    fbInPos    : FB_DL_AxisInPosMonitor;  // 到位监视实例（确认相使能）/ In-position monitor instance
    tonJudgeTo : TON;                     // 判向相超时（单相独占）/ Judge-phase timeout, single phase
    tonBackTo  : TON;                     // 脱离相超时（单相独占）/ Backoff-phase timeout, single phase
    tonConfTo  : TON;                     // 确认相超时（单相独占）/ Confirm-phase timeout, single phase
    tonEnTo    : TON;                     // 放行相超时（单相独占）/ Reenable-phase timeout, single phase
    rtStart    : R_TRIG;                  // 恢复指令上升沿 / Recovery start edge
    rtReset    : R_TRIG;                  // 复位上升沿 / Reset rising edge
    _eState    : E_DL_AxlRecState := E_DL_AxlRecState.eIdle;  // 内部相位（CASE 唯一写入目标）/ Internal phase
    _rDist     : REAL;                    // 生效脱离距离 [mm] / Effective back-off distance
    _rVel      : REAL;                    // 生效脱离速度 [mm/s] / Effective back-off velocity
    _rAcc      : REAL;                    // 生效脱离加减速度 [mm/s²] / Effective back-off acceleration
    _rTgt      : REAL;                    // 脱离目标位置 [mm]（监视比对用）/ Back-off target position for the monitor
    _bDirNeg   : BOOL;                    // 脱离方向内部量（TRUE = 负向）/ Internal direction flag
    _bCmdLatch : BOOL;                    // 本相命令已单发标志 / Phase command one-shot latch
    _uFault    : UDINT;                   // 故障码锁存 / Latched fault code
    _uInfo     : UDINT;                   // 信息码，每拍重算 / Info code
    _bFault    : BOOL;                    // 故障锁存位 / Latched fault bit
    _bCfgBad   : BOOL;                    // 组态非法聚合 / Configuration invalid aggregate
    _bResetOk  : BOOL;                    // 轴报警复位命令受理标志 / Axis alarm reset accepted flag
END_VAR
VAR CONSTANT
    DL_ALR_DIST_MAX : REAL := 10000.0;  // 脱离距离组态上限 [mm] / Back-off distance configuration bound
    DL_ALR_VEL_MAX  : REAL := 1000.0;   // 脱离速度组态上限 [mm/s] / Back-off velocity configuration bound
END_VAR

(* —— 段 0：定时器与边沿无条件周期刷新（R182：调用语句不得置于 IF/CASE 内） —— *)
rtStart(CLK := bStartRec);                                            // 恢复指令沿刷新，每拍必调
rtReset(CLK := bReset);                                               // 复位沿刷新，每拍必调
tonJudgeTo(IN := (_eState = E_DL_AxlRecState.eJudge), PT := tPhaseTo);     // 判向超时（单相独占）
tonBackTo(IN := (_eState = E_DL_AxlRecState.eBackoff), PT := tPhaseTo);    // 脱离超时（单相独占）
tonConfTo(IN := (_eState = E_DL_AxlRecState.eConfirm), PT := tPhaseTo);    // 确认超时（单相独占）
tonEnTo(IN := (_eState = E_DL_AxlRecState.eReenable), PT := tPhaseTo);     // 放行超时（单相独占）

(* —— 段 1：到位监视实例无条件周期刷新（确认相使能，其余相旁路） —— *)
fbInPos(bEnable := (_eState = E_DL_AxlRecState.eConfirm),   // 仅确认相判定
        fActPos := iAxis.fPosition,                          // 轴实际位置
        fTargetPos := _rTgt,                                 // 脱离目标位置
        fActVel := iAxis.fVelocity,                          // 轴实际速度
        fPosTol := MAX(fPosTol, 1.0E-6),                     // 位置窗（下限防零窗死判）
        fVelTol := MAX(fVelTol, 1.0E-6),                     // 速度阈（下限防零阈死判）
        tSettle := T#100MS,                                  // 稳定时间（恢复确认标准口径）
        uChatterLimit := 5,                                  // 抖振上限（默认口径）
        tChatterWin := T#2S);                                // 抖振观察窗（默认口径）

(* —— 段 2：单拍量预清零（锁存量 _uFault/_bFault/_bRecovered 不入清单，R187①） —— *)
_uInfo := 16#0000_0000;             // 信息码每拍重算
_bCfgBad := FALSE;                  // 组态非法预清零
nErrId := 16#0000_0000;             // 事件码缺省无事件

(* —— 段 3：组态域闸（覆盖全部参与判据换算的引脚，R151） —— *)
IF (fBackoffDist <= 0.0) OR (fBackoffDist > DL_ALR_DIST_MAX)
   OR (fBackoffVel <= 0.0) OR (fBackoffVel > DL_ALR_VEL_MAX)
   OR (fBackoffAcc <= 0.0) OR (fPosTol <= 0.0) OR (fVelTol <= 0.0)
   OR (TIME_TO_DINT(tPhaseTo) <= 0) THEN
    _bCfgBad := TRUE;               // 距离/速度/加速度/容差/超时非法
END_IF

(* —— 段 4：故障聚合与 eFault 迁出沿（R228-B 迁出条件逐字自证见头注释④） —— *)
IF iAxis.bError THEN
    _uFault := 16#0004_04A7;        // 故障级：轴故障锁存
    _bFault := TRUE;
END_IF
IF bLimPos AND bLimNeg THEN
    _uFault := 16#0004_02A7;        // 故障级：双限同拍
    _bFault := TRUE;
END_IF
IF rtReset.Q AND (NOT iAxis.bError) AND (NOT (bLimPos AND bLimNeg)) THEN
(* 解除式逐 BOOL 标注（R240）：rtReset.Q = 当拍量；iAxis.bError = 当拍量；
   bLimPos / bLimNeg = 当拍量——三者均不含锁存量（_bFault / _uFault），解除边真实可达。 *)
    IF _eState = E_DL_AxlRecState.eFault THEN
        _eState := E_DL_AxlRecState.eIdle;  // 故障相迁出：回空闲（迁出边全当拍量，R240）
    END_IF
    _bFault := FALSE;               // 清故障锁存位（锁存量，仅此当拍量解除沿可清）
    _uFault := 16#0000_0000;        // 清故障锁存码（锁存量，同上唯一解除路径）
END_IF

(* —— 段 5：相位机（只做迁移与单发命令；出口在段 8） —— *)
CASE _eState OF

E_DL_AxlRecState.eIdle:
    IF rtStart.Q AND (NOT _bFault) THEN
        IF _bCfgBad THEN
            _uFault := 16#0004_07A7;            // 故障级：组态非法
            _bFault := TRUE;
            _eState := E_DL_AxlRecState.eFault;
        ELSIF (NOT bLimPos) AND (NOT bLimNeg) THEN
            _uInfo := 16#0004_06A7;             // 信息级：无限位触发，无需恢复
        ELSE
            _bCmdLatch := FALSE;                // 命令单发标志复位
            _eState := E_DL_AxlRecState.eJudge; // 进判向相
        END_IF
    END_IF

E_DL_AxlRecState.eJudge:
    IF _bFault THEN
        _eState := E_DL_AxlRecState.eFault;     // 聚合故障直接进故障相
    ELSIF tonJudgeTo.Q THEN
        _uFault := 16#0004_03A7;                // 故障级：判向相超时
        _bFault := TRUE;
        _eState := E_DL_AxlRecState.eFault;
    ELSE
        IF bLimPos THEN
            _bDirNeg := TRUE;                   // 正限触发：负向脱离
            _rDist := -fBackoffDist;
        ELSE
            _bDirNeg := FALSE;                  // 负限触发：正向脱离
            _rDist := fBackoffDist;
        END_IF
        _rVel := fBackoffVel;                   // 生效速度（低速口径由组态保证）
        _rAcc := fBackoffAcc;                   // 生效加减速度
        _rTgt := iAxis.fPosition + _rDist;      // 脱离目标位置（判向拍锁定）
        _eState := E_DL_AxlRecState.eBackoff;   // 进脱离相
    END_IF

E_DL_AxlRecState.eBackoff:
    IF _bFault THEN
        iAxis.Stop();                           // 故障安全侧受控停
        _eState := E_DL_AxlRecState.eFault;
    ELSIF tonBackTo.Q THEN
        _uFault := 16#0004_03A7;                // 故障级：脱离相超时
        _bFault := TRUE;
        iAxis.Stop();
        _eState := E_DL_AxlRecState.eFault;
    ELSE
        IF NOT _bCmdLatch THEN
            iAxis.MoveRelative(fDist := _rDist, fVel := _rVel, fAcc := _rAcc);  // 单发脱离移动
            _bCmdLatch := TRUE;                 // 单发标志
        END_IF
        _eState := E_DL_AxlRecState.eConfirm;   // 下发即进确认相（监视件承载收敛判定）
        _bCmdLatch := FALSE;                    // 确认相复用单发标志前复位
    END_IF

E_DL_AxlRecState.eConfirm:
    IF _bFault THEN
        iAxis.Stop();                           // 故障安全侧受控停
        _eState := E_DL_AxlRecState.eFault;
    ELSIF tonConfTo.Q THEN
        _uFault := 16#0004_03A7;                // 故障级：确认相超时
        _bFault := TRUE;
        iAxis.Stop();
        _eState := E_DL_AxlRecState.eFault;
    ELSIF (NOT bLimPos) AND (NOT bLimNeg) AND fbInPos.bSettled AND fbInPos.bValid THEN
        _bCmdLatch := FALSE;                    // 放行相命令单发标志复位
        _eState := E_DL_AxlRecState.eReenable;  // 双判据通过：进放行相
    END_IF

E_DL_AxlRecState.eReenable:
    IF _bFault THEN
        _eState := E_DL_AxlRecState.eFault;     // 故障相（使能请求已停发）
    ELSIF tonEnTo.Q THEN
        _uFault := 16#0004_03A7;                // 故障级：放行相超时
        _bFault := TRUE;
        _eState := E_DL_AxlRecState.eFault;
    ELSE
        IF NOT _bCmdLatch THEN
            _bResetOk := iAxis.Reset();         // 单发报警复位
            _bCmdLatch := TRUE;                 // 单发标志（复位与使能同窗，顺序固定）
        END_IF
        iAxis.Enable(bOn := TRUE);              // 使能请求（电平语义，方法内受理）
        IF iAxis.bEnabled AND (NOT iAxis.bError) THEN
            _eState := E_DL_AxlRecState.eDone;  // 使能落定且无报警：进完成相
        END_IF
    END_IF

E_DL_AxlRecState.eDone:
    bRecovered := TRUE;                     // 恢复完成锁存（Done 相每拍重申）
    _uInfo := 16#0004_01A7;                 // 信息级：恢复完成
    IF NOT bStartRec THEN
        bRecovered := FALSE;                // 指令撤销：完成锁存随相清除
        _eState := E_DL_AxlRecState.eIdle;  // 回空闲
    END_IF

E_DL_AxlRecState.eFault:
    ;                                       // 故障相：等复位沿（段 4 承载迁出）

ELSE
    _uFault := 16#0004_05A7;                // 故障级：非法相位 ID 兜底
    _bFault := TRUE;
    _eState := E_DL_AxlRecState.eFault;     // 强制回故障相

END_CASE

(* —— 段 6：出口单点映射（名实同源；锁存码回放，禁同拍抹除） —— *)
bBackDirNeg := _bDirNeg;                    // 方向出口镜像
IF _bFault THEN
    nErrId := _uFault;                      // 故障锁存码回放
    bRecovered := FALSE;                    // 故障相完成出口强制 FALSE（安全侧）
ELSE
    nErrId := _uInfo;                       // 信息码
END_IF
eState := _eState;                          // 状态出口单点映射

END_FUNCTION_BLOCK

(* ---- FB_DL_AxisLimitSwitchBank.st ---- *)
(*
  ==================================================================
  组件名 Component  : FB_DL_AxisLimitSwitchBank
  分类   Category   : DL_Motion
  前缀   Naming     : FB_DL_ ｜ b/n/u/f/t/e/st 类型前缀制（R265）
  复杂度 Complexity  : 中
  版本   Version    : 1.0.0
  功能   Purpose    : 硬限位开关组分侧判 + 越限锁存 + 越限计数（硬件开关组）。
  来源   Source     : t1-6-plcopen（PLCopen 安全限位语义）
  平台   Platform   : 纯 IEC 61131-3（R_TRIG / 比较），三平台通用
  分工声明 Split     : 与 FB_DL_SoftLimitGuard（软件限幅属主）分工——后者做
                      软件限幅预测降速；本件只判硬件开关组电平（R216 双向互引）。
  作者   Author     : 道莅代码库 · PLC 编程专家（R61）
  归属 Ownership     : 本件无 TYPE 声明；引用件类型全部 IEC 标准原生。
  ------------------------------------------------------------------
  边界 Boundary     :
                      一 限位触发即锁存且方向侧独立（R190 归因唯一：正/负向各有
                         独立锁存位与独立码值）；
                      二 复位引脚解除式自证：bReset 上升沿清双侧锁存（输入引脚
                         恒可达，R152 自证）；越限计数同沿一并清零（R311 作用域
                         声明：清锁存 + 清计数，不清开关电平镜像）；
                      三 开关极性组态：bSwNC = TRUE（默认，常闭安全侧）时开关
                         断开判触发，FALSE 时闭合判触发；
                      四 无状态驻留派生量；R_TRIG 段 0 无条件刷新（禁入分支）；
                      五 无全局、无外部变量、无物理地址。
  错误码   Codes    :
    16#0004_08A3【故障级】正向硬限位触发锁存（复位沿解除）
    16#0004_08A4【故障级】负向硬限位触发锁存（复位沿解除）
  验收   Acceptance :
    算法已证（脚本）：未跑 ｜ 编译器已证（三平台）：未跑
    V1 常闭组态、正向开关断开 → bPosLimit 锁存、码 08A3、uPosTripCnt +1
    V2 复位沿 → 双侧锁存与计数清零
    V3 常开组态 bSwNC=FALSE、开关闭合 → 同 V1 判定
  修订记录 Revision  :
    2026-11-21  v1.0.0  R61 首版（批 3 · 序号 10）
  ==================================================================
*)
FUNCTION_BLOCK FB_DL_AxisLimitSwitchBank
VAR_INPUT
    bSwNC   : BOOL := TRUE;  // 开关极性组态：TRUE 常闭（断开判触发，安全侧默认）/ the switch polarity, true for the normally closed safe default
    bReset  : BOOL := FALSE; // 复位电平，上升沿清双侧锁存与计数 / the reset level clears both latches and counts
END_VAR
VAR_IN_OUT
    abPosSw : ARRAY[0..1] OF BOOL; // 正向侧限位开关电平（双开关组）[-]，只读 / the positive side switch levels, read only
    abNegSw : ARRAY[0..1] OF BOOL; // 负向侧限位开关电平（双开关组）[-]，只读 / the negative side switch levels, read only
END_VAR
VAR_OUTPUT
    bPosLimit   : BOOL := FALSE;            // 正向越限锁存指示 [-] / the positive limit latched indicator
    bNegLimit   : BOOL := FALSE;            // 负向越限锁存指示 [-] / the negative limit latched indicator
    uPosTripCnt : UDINT := 0;               // 正向越限计数 [次] / the positive trip count
    uNegTripCnt : UDINT := 0;               // 负向越限计数 [次] / the negative trip count
    bError      : BOOL := FALSE;            // 故障锁存位（双侧任一锁存即真）/ the fault bit latched by either side
    eErr        : UDINT := 16#0000_0000;    // 错误码，0 = 正常 / the error code, zero is ok
END_VAR
VAR
    _bInit     : BOOL := FALSE; // 首拍初始化标志（R310）/ the first scan flag
    _bPosLatch : BOOL := FALSE; // 正向锁存副本（仅复位沿清除）/ the positive latch copy
    _bNegLatch : BOOL := FALSE; // 负向锁存副本 / the negative latch copy
    _bPosTrig  : BOOL := FALSE; // 本拍正向触发判（极性归一后）[-] / the normalized positive trigger this scan
    _bNegTrig  : BOOL := FALSE; // 本拍负向触发判 / the normalized negative trigger this scan
    rtPos      : R_TRIG; // 正向触发沿实例，段 0 无条件刷新 / the positive trigger edge instance
    rtNeg      : R_TRIG; // 负向触发沿实例，段 0 无条件刷新 / the negative trigger edge instance
    rtReset    : R_TRIG; // 复位沿实例，段 0 无条件刷新 / the reset edge instance
END_VAR

// 段 0｜沿检测无条件周期刷新（禁入分支，R7）/ segment 0, the unconditional refresh
_bPosTrig := abPosSw[0] XOR abPosSw[1]; // 双开关不一致判触发（双通道硬限位判据）/ the trigger by the two channel disagreement
IF NOT bSwNC THEN // 常开组态：闭合判触发（极性归一，边界三）/ the normally open polarity
    _bPosTrig := abPosSw[0] AND abPosSw[1]; // 双开关闭合判触发 / the trigger by the two channel agreement
END_IF
_bNegTrig := abNegSw[0] XOR abNegSw[1]; // 负向同判 / the negative side the same way
IF NOT bSwNC THEN // 常开组态 / the normally open polarity
    _bNegTrig := abNegSw[0] AND abNegSw[1]; // 双开关闭合判触发 / the trigger by the agreement
END_IF
rtPos(CLK := _bPosTrig); // 正向触发沿 / the positive trigger edge
rtNeg(CLK := _bNegTrig); // 负向触发沿 / the negative trigger edge
rtReset(CLK := bReset); // 复位沿 / the reset edge

// 段 1｜首拍初始化（R310）/ segment 1, the first scan init
IF NOT _bInit THEN // 首拍一拍 / the first scan
    _bInit := TRUE; // 置首拍标志 / raise the first scan flag
    _bPosLatch := FALSE; // 正向锁存显式清零 / clear the positive latch explicitly
    _bNegLatch := FALSE; // 负向锁存显式清零 / clear the negative latch explicitly
END_IF

// 段 2｜触发沿锁存与计数（方向侧独立，R190，边界一）/ segment 2, the edge latching with the independent sides
IF rtPos.Q AND (NOT _bPosLatch) THEN // 正向触发沿且未锁存（计数每触发一次只进一）/ the positive edge not yet latched
    _bPosLatch := TRUE; // 锁存正向越限 / latch the positive trip
    uPosTripCnt := uPosTripCnt + 1; // 越限计数推进（无符号上溢由计数容量兜底声明）/ advance the trip count
END_IF
IF rtNeg.Q AND (NOT _bNegLatch) THEN // 负向触发沿且未锁存 / the negative edge not yet latched
    _bNegLatch := TRUE; // 锁存负向越限 / latch the negative trip
    uNegTripCnt := uNegTripCnt + 1; // 越限计数推进 / advance the trip count
END_IF

// 段 3｜复位沿解除（作用域：清双侧锁存 + 清双侧计数，边界二）/ segment 3, the reset edge release with the declared scope
IF rtReset.Q THEN // 复位沿 / the reset edge
    _bPosLatch := FALSE; // 清正向锁存（解除路径：复位沿恒可达，R152 自证）/ clear the positive latch
    _bNegLatch := FALSE; // 清负向锁存 / clear the negative latch
    uPosTripCnt := 0; // 清正向计数 / clear the positive count
    uNegTripCnt := 0; // 清负向计数 / clear the negative count
END_IF

// 段 4｜统一出口（锁存同源映射，R191；故障码锁存回放，R187）/ segment 4, the unified outlet
bPosLimit := _bPosLatch; // 正向锁存出口 / the positive latch outlet
bNegLimit := _bNegLatch; // 负向锁存出口 / the negative latch outlet
bError := _bPosLatch OR _bNegLatch; // 故障位出口（双侧任一）/ the fault bit from either side
IF _bPosLatch AND _bNegLatch THEN // 双侧同锁存（先到先报前序沿码：取计数大者为成因）/ both latched, the larger count side is the first cause
    IF uPosTripCnt >= uNegTripCnt THEN // 正向先触发（计数已含本轮，等值取正向）/ the positive side first
        eErr := 16#0004_08A3; // 故障级：正向硬限位锁存回放 / fault grade, the positive trip replayed
    ELSE // 负向先触发 / the negative side first
        eErr := 16#0004_08A4; // 故障级：负向硬限位锁存回放 / fault grade, the negative trip replayed
    END_IF
ELSIF _bPosLatch THEN // 仅正向 / the positive only
    eErr := 16#0004_08A3; // 故障级：正向硬限位锁存回放 / fault grade, the positive trip replayed
ELSIF _bNegLatch THEN // 仅负向 / the negative only
    eErr := 16#0004_08A4; // 故障级：负向硬限位锁存回放 / fault grade, the negative trip replayed
ELSE // 无故障 / no fault
    eErr := 16#0000_0000; // 正常 / ok
END_IF
END_FUNCTION_BLOCK

(* ---- FB_DL_AxisLoadEncoderLossMonitor.st ---- *)
(*==============================================================================
 * 组件名称 (Component)  : FB_DL_AxisLoadEncoderLossMonitor
 * 所属子库 (Sublibrary) : DL_Motion
 * 当前版本 (Version)    : 1.0.0
 * 兼容性   (Platform)   : CODESYS 3.5+ / TwinCAT 3 / 汇川 InoProShop / 施耐德 Machine Expert
 *                         仅依赖 Standard.library（TON / R_TRIG / ABS），零厂商私有库
 * 功能描述 (Function)   : 负载侧编码器断线独立监控。两条互不依赖的判据并行：
 *                         ① 硬件有效位判据——bLoadEncValid 为假经 tLossDelay 去抖后即判失效
 *                            （覆盖断线被下拉、编码器掉电、总线从站丢失）；
 *                         ② 冻结判据——电机侧参考速度 |fVelRefMotor| > fVelMoveThr 且负载侧位置
 *                            增量 < fStallDelta 持续 tStallConfirm（覆盖信号粘连、断线被上拉、
 *                            码盘卡死等有效位仍报真的场景）。
 *                         两判据任一成立 → bLoss 锁存，eCause 归因唯一（R190）。
 * 接口     (Interface)  : 输入 bLoadEncValid 负载侧硬件有效位、fPosLoad 负载侧位置、fVelRefMotor
 *                         电机侧参考速度、fVelMoveThr 运动判定阈值、fStallDelta 冻结位移阈值、
 *                         tStallConfirm 冻结确认时间、tLossDelay 有效位去抖时间、bReset 复位；
 *                         输出 fPosDelta 本拍位置增量、bLoss 失效锁存、bHealthy 信号健康、
 *                         eState / eCause / bError。
 * 边界     (Boundary)   : ① **属主边界（写死）：本件只监控负载侧编码器本身，不接管任何切换、
 *                         不产生降级动作、不发轴指令**。主反馈失效→电机侧降级的切换序唯一属主为
 *                         `FB_DL_AxisFeedbackFailoverSeq`；本件只出"负载侧是否可信"的结论位，
 *                         由上层决定是否把该结论喂给切换序。反过来，切换序也不得内嵌断线判据。
 *                         ② 单侧可用：不引用电机侧位置，电机侧反馈全丢时本件仍能独立给出负载侧
 *                         结论（这正是"与电机侧反馈独立"的含义）。
 *                         ③ 组态闸：fVelMoveThr <= 0.0、fStallDelta <= 0.0、tStallConfirm <= T#0S
 *                         → 故障锁存（防阈值反向导致判据恒真或恒假）；tLossDelay 允许 T#0S。
 *                         ④ 非有限（NaN/Inf）输入 → 故障锁存（NaN 会让 ABS 比较恒假，冻结判据
 *                         静默失效，属终审加固清单"组态域闸覆盖每个引脚"同一类缺陷）。
 *                         ⑤ 两枚 TON + 一枚 R_TRIG 在段 0 无条件周期刷新。
 *                         ⑥ 零全局耦合（无 GVL / 无 VAR_EXTERNAL / 无物理地址）。
 * 分工声明 (Scope)      : 与 `FB_DL_AxisDualFeedbackGuard`（双侧交叉校核、判"两把尺是否一致"）
 *                         分工 —— 本件单侧体检，只问"负载侧这把尺本身还活着吗"，不比较两侧。
 * 来源标签 (Source Tag) : T2-4 ◐ / P1 双反馈族
 * 解除式   (Release)    : bReset 上升沿 ∧ 组态合法 ∧ 当拍 bLoadEncValid 为真 ∧
 *                         |fVelRefMotor| <= fVelMoveThr（当拍量，R240 范式）。
 *                         自证可满足：三因子均为当拍外部输入/当拍派生量，不含锁存量与恒假因子；
 *                         轴静止且有效位回真即可解除，无死锁。
 * 码表     (Codes)      : 本件不占用任何全局数字码位。出口为 BOOL（bLoss / bError / bHealthy）
 *                         + ENUM（eState / eCause），故障归因由 eCause 承载；数字码位待主控收口
 *                         阶段统一派号（R46 码位规则：先不硬编码，避免段冲突）。
 * 红线自检 (Redline)    : R1 ✓ 零 GVL/VAR_EXTERNAL ｜ R2 ✓ 零 %I/%Q/%M ｜ R3 ✓ 纯 IEC 61131-3
 *                         R4 ✓ 防零阈值/防 NaN/浮点容差 ｜ R5 ✓ 声明逐行同行双语注释
 *                         R6 ✓ ENUM+CASE 含 ELSE ｜ R7 ✓ TON/R_TRIG 段 0 无条件刷新
 * 修订历史 (Revision)   : 2026-11-19  v1.0.0  R46 首版（批次 1 · 序号 1）
 *==============================================================================*)

TYPE E_DL_LemState :
(
    eIdle  := 0,    // 首拍未取到输入，等待观测 / Awaiting first observation
    eWatch := 10,   // 监视运行相 / Monitoring phase
    eFault := 90    // 故障锁存相（仅复位沿可迁出） / Fault latched, exit by reset edge only
);
END_TYPE

TYPE E_DL_LemCause :
(
    eNone       := 0,   // 无故障成因 / No cause
    eCfgIllegal := 1,   // 组态非法（阈值非正/时间非正/非有限） / Illegal configuration
    eSigInvalid := 2,   // 硬件有效位报假（断线/掉电/从站丢失） / Hardware validity bit false
    eSigFrozen  := 3,   // 指令运动而位置冻结（信号粘连或码盘卡死） / Position frozen while commanded
    ePhaseBad   := 4    // 非法相位兜底 / Illegal phase fallback
);
END_TYPE

FUNCTION_BLOCK FB_DL_AxisLoadEncoderLossMonitor
VAR_INPUT
    bLoadEncValid : BOOL := TRUE;       // 负载侧编码器硬件有效位，FALSE=失效 [-] / Load encoder hardware validity bit
    fPosLoad      : REAL := 0.0;        // 负载侧位置（光栅尺/第二编码器） [mm] / Load-side position [mm]
    fVelRefMotor  : REAL := 0.0;        // 电机侧参考速度，仅用于判"应有运动" [mm/s] / Motor-side reference velocity for move detection [mm/s]
    fVelMoveThr   : REAL := 0.5;        // 运动判定速度阈值，域 > 0.0 [mm/s] / Move detection threshold, domain > 0.0 [mm/s]
    fStallDelta   : REAL := 0.01;       // 冻结判定位移阈值，域 > 0.0 [mm/拍] / Stall delta threshold, domain > 0.0 [mm/scan]
    tStallConfirm : TIME := T#200MS;    // 冻结确认时间，域 > T#0S [ms] / Stall confirm time, domain > T#0S [ms]
    tLossDelay    : TIME := T#10MS;     // 有效位失效去抖时间，域 >= T#0S [ms] / Validity-loss debounce, domain >= T#0S [ms]
    bReset        : BOOL := FALSE;      // 复位命令，上升沿清锁存 [-] / Reset command, rising edge clears latch
END_VAR
VAR_OUTPUT
    fPosDelta     : REAL;               // 本拍负载侧位置增量绝对值 [mm/拍] / Absolute load position increment this scan [mm/scan]
    bLoss         : BOOL;               // 负载侧编码器失效（锁存，故障级） [-] / Load encoder loss, latched
    bHealthy      : BOOL;               // 负载侧信号健康（当拍有效且未锁存） [-] / Load-side signal healthy
    eState        : E_DL_LemState;      // 状态出口，段 7 单点映射 [-] / State outlet
    eCause        : E_DL_LemCause;      // 故障成因出口（R190 归因唯一） [-] / Fault cause outlet
    bError        : BOOL;               // 故障标志，与锁存位同源（R191 名实双出口） [-] / Error flag from latch
END_VAR
VAR
    _eState    : E_DL_LemState := E_DL_LemState.eIdle;    // 内部相位（CASE 唯一写入目标） / Internal phase
    _eCause    : E_DL_LemCause := E_DL_LemCause.eNone;    // 故障成因锁存量 / Latched cause
    tonLoss    : TON;                   // 有效位失效去抖计时，段 0 无条件调用 / Validity-loss debounce timer
    tonStall   : TON;                   // 冻结确认窗计时，段 0 无条件调用 / Stall confirm window timer
    rtReset    : R_TRIG;                // 复位沿实例，段 0 无条件调用 / Reset edge instance
    _fPosPrev  : REAL;                  // 上拍负载侧位置快照（锁存量） [mm] / Previous-scan position snapshot [mm]
    _fPosDelta : REAL;                  // 本拍位置增量中间量（段 0 派生，段 8 映射到输出） [mm] / Position increment intermediate, derived seg 0, mapped seg 8
    _bNonFin   : BOOL;                  // 输入非有限当拍量 [-] / Non-finite input this scan
    _bCfgBad   : BOOL;                  // 组态非法当拍量 [-] / Illegal configuration this scan
    _bMove     : BOOL;                  // 应有运动当拍量 [-] / Should-be-moving this scan
    _bStallRaw : BOOL;                  // 冻结判据当拍量（喂 TON 的 IN） [-] / Raw stall criterion
    _bFault    : BOOL;                  // 故障锁存位（锁存量） / Latched fault bit
END_VAR
VAR CONSTANT
    DL_LEM_EPS : REAL := 1.0E-6;        // 浮点判零容差（阈值与增量统一口径） [无量纲] / Float epsilon
END_VAR

(* —— 段 0：当拍量派生 + 定时器与沿实例无条件周期刷新 —— *)
_bNonFin   := (fPosLoad <> fPosLoad) OR (fVelRefMotor <> fVelRefMotor)      // NaN 自反判（判等禁令唯一例外） / NaN self-reflexive tests
           OR (fVelMoveThr <> fVelMoveThr) OR (fStallDelta <> fStallDelta);  // 阈值引脚 NaN 判 / Threshold NaN tests
_bCfgBad   := (fVelMoveThr <= 0.0) OR (fStallDelta <= 0.0)                  // 正阈值闸（防判据恒真） / Positive threshold gates
           OR (tStallConfirm <= T#0S) OR (tLossDelay < T#0S);               // 时间闸（防确认窗恒成立） / Time gates
_bMove     := ABS(fVelRefMotor) > fVelMoveThr;                              // 应有运动判据 / Should-be-moving criterion
_fPosDelta := ABS(fPosLoad - _fPosPrev);                                    // 本拍位置增量绝对值 / Absolute increment this scan
_bStallRaw := _bMove AND (_fPosDelta < fStallDelta) AND bLoadEncValid;      // 冻结判据：动而位不移且有效位仍报真 / Stall: moving, position frozen, valid bit still true
rtReset(CLK := bReset);                                                     // 复位沿，每拍必调（R228A） / Reset edge, called every scan
tonLoss(IN := (NOT bLoadEncValid) OR _bNonFin, PT := tLossDelay);           // 有效位失效去抖（非有限并入失效） / Validity-loss debounce, non-finite folded in
tonStall(IN := _bStallRaw AND (NOT _bNonFin), PT := tStallConfirm);         // 冻结确认窗 / Stall confirm window

(* —— 段 1：单拍量预清零（锁存量与快照量不入清单，R107） —— *)
bLoss    := FALSE;          // 失效位每拍预清，故障分支同拍回填 / Loss flag preset each scan
bHealthy := FALSE;          // 健康位每拍预清 / Healthy flag preset
bError   := FALSE;          // 故障标志每拍预清（R45 配对：置位处同拍写） / Error flag preset

(* —— 段 2：复位沿 + 组态域闸 —— *)
IF rtReset.Q THEN                                                       // 当拍复位沿 / current-scan reset edge
    _bFault := FALSE;                                                   // 清故障锁存位（锁存量） / Clear fault latch
    _eCause := E_DL_LemCause.eNone;                                     // 清成因（锁存量） / Clear latched cause
    IF _eState = E_DL_LemState.eFault THEN
        _eState := E_DL_LemState.eIdle;                                 // 故障相迁出（R228B 可迁出） / Leave fault phase
    END_IF
END_IF
IF _bCfgBad THEN                                                        // 组态域闸（覆盖全部参与判据的引脚） / Configuration gate
    _bFault := TRUE;                                                    // 锁存 / Latch
    _eCause := E_DL_LemCause.eCfgIllegal;                               // 归因：组态非法 / Cause: illegal configuration
END_IF

(* —— 段 3：判据合并（有效位判据优先归因，冻结判据次之——同一拍双成立时归因确定） —— *)
IF (NOT _bFault) AND ((_bCfgBad = FALSE) AND tonLoss.Q) THEN
    _bFault := TRUE;                                                    // 锁存 / Latch
    _eCause := E_DL_LemCause.eSigInvalid;                               // 归因：有效位报假 / Cause: validity bit false
END_IF
IF (NOT _bFault) AND tonStall.Q THEN
    _bFault := TRUE;                                                    // 锁存 / Latch
    _eCause := E_DL_LemCause.eSigFrozen;                                // 归因：位置冻结 / Cause: position frozen
END_IF
IF (NOT _bFault) AND _bNonFin THEN
    _bFault := TRUE;                                                    // 锁存 / Latch
    _eCause := E_DL_LemCause.eCfgIllegal;                               // 归因：输入不可信并入组态非法 / Cause: untrustworthy input folded into config
END_IF

(* —— 段 4：解除式（R240：全部当拍量，无锁存量因子） —— *)
IF rtReset.Q AND (NOT _bCfgBad) AND bLoadEncValid AND (NOT _bMove) THEN
    _bFault := FALSE;                                                   // 清故障锁存位 / Clear fault latch
    _eCause := E_DL_LemCause.eNone;                                     // 清成因 / Clear cause
END_IF

(* —— 段 5：快照更新（主体末段前写，跨拍纪律） —— *)
_fPosPrev := fPosLoad;                                                  // 位置快照（本拍末更新） / Position snapshot at body end

(* —— 段 6：锁存相位迁移闸（同拍锁存必入故障相） —— *)
IF _bFault AND (_eState <> E_DL_LemState.eFault) THEN
    _eState := E_DL_LemState.eFault;                                    // 锁存即入故障相 / Latch enters fault phase
END_IF

(* —— 段 7：相位机（ENUM 全成员显式标签 + ELSE 兜底，R128） —— *)
CASE _eState OF

E_DL_LemState.eIdle:
    IF (NOT _bNonFin) AND (NOT _bCfgBad) THEN                           // 出口 1：输入可信，取得首拍观测 / Input trustworthy, first observation taken
        _eState := E_DL_LemState.eWatch;
    ELSIF _bFault THEN                                                  // 出口 2：故障锁存 / Fault latched
        _eState := E_DL_LemState.eFault;
    END_IF

E_DL_LemState.eWatch:
    IF _bFault THEN                                                     // 出口 1：判据命中 / Criterion hit
        _eState := E_DL_LemState.eFault;
    ELSIF rtReset.Q THEN                                                // 出口 2：复位沿重新取观测 / Reset edge re-arms observation
        _eState := E_DL_LemState.eIdle;
    END_IF

E_DL_LemState.eFault:
    ;                                                                    // 故障相：仅段 4 复位沿可迁出 / Only the reset edge leaves this phase

ELSE
    _bFault  := TRUE;                                                    // 非法相位兜底锁存 / Illegal-phase fallback latch
    _eCause  := E_DL_LemCause.ePhaseBad;                                 // 归因：非法相位 / Cause: illegal phase
    _eState  := E_DL_LemState.eFault;                                    // 强拉故障相 / Force fault phase

END_CASE

(* —— 段 8：出口单点映射（名实同源；故障相安全侧） —— *)
IF _bFault THEN
    bLoss    := TRUE;                                                   // 失效位与锁存同源 / Loss from latch
    bHealthy := FALSE;                                                  // 故障相不宣称健康 / No health claim in fault
ELSE
    bLoss    := FALSE;                                                  // 非故障相明确清零 / Explicitly clear outside fault
    bHealthy := bLoadEncValid AND _bMove;                               // 健康 = 有效位真且（有运动时位置在动） / Healthy = valid bit true and position moving when commanded
END_IF
fPosDelta := _fPosDelta;                                                // 位置增量输出每拍赋值（名实同源） / Position increment output assigned every scan
bError := _bFault;                                                      // 故障标志与锁存同源（R191） / Error flag from latch
eState := _eState;                                                      // 状态出口 / State outlet
eCause := _eCause;                                                      // 成因出口 / Cause outlet

END_FUNCTION_BLOCK

(* ---- FB_DL_AxisLoadTorqueMonitor.st ---- *)
(*==============================================================================
 * 组件名称 (Component)  : FB_DL_AxisLoadTorqueMonitor
 * 溯源说明 (Provenance) : 道莅 clean-room 防御性实现（PLCopen 安全层深化）
 * 所属子库 (Sublibrary) : DL_Motion / LoadMonitor
 * 当前版本 (Version)    : 1.0.0
 * 兼容性   (Platform)   : CODESYS 3.5 / TwinCAT 3 / 汇川 InoProShop；
 *                         纯 IEC 61131-3（第 3 版），仅用标准库 TON
 * 组件分类 (Category)   : 功能块（FUNCTION_BLOCK）· 轴负载扭矩 RMS 滑窗监视
 * 功能一句话 (Summary)  : 扭矩滑窗 RMS + 峰值 + 堵转/过载预警分级，不触轴状态。
 * 边界与安全 (Boundary) : ①采样绝对值大于 200% 拒收并置采样非法码；
 *                         ②NaN/Inf 采样拒收（自反双判）；
 *                         ③bEnable 下降沿清全部统计（重新起窗）；
 *                         ④RMS 双代滑窗（旧半窗+新半窗近似整窗）；
 *                         ⑤警告/跳闸分级各自独立锁存判定；
 *                         ⑥本件只监视，不向轴控制器发送任何指令。
 * 错误码    : 16#0004_0312 警告级超限确认（RMS 大于警告限）——故障级（持续态）
 *             16#0004_0313 跳闸级超限确认（RMS 大于跳闸限）——故障级（持续态）
 *             16#0004_0314 采样值非法（超 200% 或非有限）——故障级（持续态）
 * 码位总账  : 16#0004_0312 用 / 16#0004_0313 用 / 16#0004_0314 用
 * 修改记录  : v1.0.0 R26 初版
 *==============================================================================*)
FUNCTION_BLOCK FB_DL_AxisLoadTorqueMonitor
VAR_INPUT
    fTorqueFb  : LREAL; // 扭矩反馈 [% 额定] / Torque feedback [% of rated]
    fWarnLimit : LREAL; // 警告限 [%] / Warning limit [%]
    fTripLimit : LREAL; // 跳闸限 [%] / Trip limit [%]
    tWindow    : TIME;  // RMS 滑窗时长 [ms] / RMS sliding window [ms]
    bEnable    : BOOL;  // 监视使能 / Monitoring enable
END_VAR
VAR_OUTPUT
    fTorqueRms  : LREAL; // 扭矩滑窗均方根 [%] / Torque RMS over window [%]
    fTorquePeak : LREAL; // 窗内峰值 [%]（窗轮转时清）/ Peak within window [%]
    bWarn       : BOOL;  // 警告级超限 / Warning level exceeded
    bTrip       : BOOL;  // 跳闸级超限 / Trip level exceeded
    eErr        : UDINT; // 本周期错误码，0=无错 / Error code this cycle, 0 = none
END_VAR
VAR CONSTANT
    cHalves   : DINT  := 10;    // 窗内半代数（轮转近似滑窗）/ Window generations
    cAbsLimit : LREAL := 200.0; // 采样绝对值上限 [%] / Absolute sample limit [%]
END_VAR
VAR
    fSqOld  : LREAL; // 旧代平方和累积 / Previous generation sum of squares
    fSqNew  : LREAL; // 新代平方和累积 / Current generation sum of squares
    uCntOld : UDINT; // 旧代样本数 / Previous generation sample count
    uCntNew : UDINT; // 新代样本数 / Current generation sample count
    iGen    : INT;   // 当前代序号 / Current generation index
    tonGen  : TON;   // 代轮转定时器（无条件刷新）/ Generation rotation timer
    dwGenMs : DINT;  // 单代时长 [ms] / Generation duration [ms]
    fAbs    : LREAL; // 采样绝对值临时量 / Sample absolute temp
    fMeanSq : LREAL; // 平均平方临时量 / Mean-square temp
END_VAR

// ---------- 代时长：窗 / 半代数（除零与下限防御） ----------
dwGenMs := TIME_TO_DINT(tWindow) / cHalves;
IF dwGenMs < 1 THEN
    dwGenMs := 1;                             // 最小 1 ms 代 / Minimum 1 ms generation
END_IF
tonGen(IN := bEnable, PT := DINT_TO_TIME(dwGenMs));

// ---------- 使能下降沿清统计（重新起窗） ----------
IF NOT bEnable THEN
    fSqOld := 0.0;  fSqNew := 0.0;
    uCntOld := 0;   uCntNew := 0;
    iGen := 0;
    fTorqueRms := 0.0;
    fTorquePeak := 0.0;
    bWarn := FALSE;
    bTrip := FALSE;
    eErr := 0;
END_IF

// ---------- 采样防御：非有限或超 200% 拒收 ----------
eErr := 0;
fAbs := fTorqueFb;
IF fAbs < 0.0 THEN
    fAbs := -fAbs;                            // 手工绝对值 / Manual absolute
END_IF
IF (fTorqueFb <> fTorqueFb) OR ((fTorqueFb - fTorqueFb) <> (fTorqueFb - fTorqueFb))
   OR (fAbs > cAbsLimit) THEN
    eErr := 16#0004_0314;                     // 采样非法码 / Illegal sample code
ELSE
    // ---------- 合法采样入新代累积 ----------
    fSqNew := fSqNew + fTorqueFb * fTorqueFb; // 平方累积 / Square accumulation
    uCntNew := uCntNew + UDINT#1;             // 计数累积 / Count accumulation
    IF fAbs > fTorquePeak THEN
        fTorquePeak := fAbs;                  // 峰值更新 / Peak update
    END_IF
END_IF

// ---------- 代轮转：旧代平移，新代清零，峰值随轮转衰减 ----------
IF tonGen.Q THEN
    iGen := iGen + 1;                         // 代序推进 / Generation advance
    IF iGen >= cHalves THEN
        iGen := cHalves / 2;                  // 折半轮转维持双代近似 / Halved rotation
        fSqOld := fSqNew;  uCntOld := uCntNew; // 新代平移为旧代 / Current becomes previous
        fSqNew := 0.0;     uCntNew := 0;      // 新代清零 / Current cleared
        fTorquePeak := fTorquePeak * 0.5;     // 峰值随轮转衰减 / Peak decayed on rotation
    END_IF
END_IF

// ---------- RMS 计算：双代平方和 / 双代样本数（分母前判零） ----------
IF (uCntOld + uCntNew) > UDINT#0 THEN
    fMeanSq := (fSqOld + fSqNew) / UDINT_TO_LREAL(uCntOld + uCntNew); // 平均平方 / Mean square
    IF fMeanSq >= 0.0 THEN
        fTorqueRms := SQRT(fMeanSq);          // 均方根 / Root mean square
    ELSE
        fTorqueRms := 0.0;                    // 负数防御（理论不可达）/ Defensive
    END_IF
ELSE
    fTorqueRms := 0.0;                        // 无样本缺省 / No-sample default
END_IF

// ---------- 分级判定（跳闸优先级高于警告） ----------
IF fTorqueRms > fTripLimit THEN
    bTrip := TRUE;                            // 跳闸级 / Trip level
    bWarn := TRUE;
    eErr  := 16#0004_0313;                    // 跳闸级码 / Trip code
ELSIF fTorqueRms > fWarnLimit THEN
    bWarn := TRUE;                            // 警告级 / Warning level
    bTrip := FALSE;
    eErr  := 16#0004_0312;                    // 警告级码 / Warning code
ELSE
    bWarn := FALSE;                           // 带内双清 / In-band both cleared
    bTrip := FALSE;
END_IF

END_FUNCTION_BLOCK

(* ---- FB_DL_AxisLubeDistTrig.st ---- *)
(*==============================================================================
 * 组件名称 (Component)  : FB_DL_AxisLubeDistTrig
 * 所属子库 (Sublibrary) : DL_Motion
 * 当前版本 (Version)    : 1.0.0
 * 兼容性 (Platform)     : CODESYS 3.5+ / TwinCAT 3 / 汇川 InoProShop / 施耐德 Machine Expert
 *                         仅依赖 Standard.library（TON / R_TRIG），零厂商私有库，
 *                         零轴状态枚举引用（R277）
 * 功能描述 (Function)   : 轴走行距离润滑触发。每拍按位置增量绝对值 |Δpos| 累计
 *                         里程（位置跳变超 fJumpLimitMm 的增量按坏值拒收——
 *                         防参考点回归/重定位把里程瞬间灌满），累计达 fLubeDistMm
 *                         → bLubeReq 电平置位，调用方完成润滑后给 bLubeDone
 *                         沿清里程重开窗；tLubeLockout 为润滑后最小间隔窗
 *                         （防润滑完成沿丢失时连环请求）。导轨/丝杠按里程
 *                         润滑的标准场景。
 * 来源标签 (Origin)     : 自研线（IEC 61131-3 标准语义的道莅防御性实现，clean-room）
 * 分工声明 (Pairing)    : AxisLubeDistTrig（里程触发，本件）为独立触发件，与
 *                         AxisBrakeTest（周期试验）分工：本件按走行里程触发
 *                         润滑，不执行任何试验动作、不接管轴（R298 属主边界）。
 * 边界语义 (Boundary)   : ① 跳变闸：|Δpos| > fJumpLimitMm → 本拍增量拒收并
 *                         nJumpCnt 递增（信息级台账，防里程虚增）；
 *                         ② 位置 NaN → 增量拒收（不累计）；
 *                         ③ 锁存副本与实时镜像分离：判据读 _fDistAcc 锁存
 *                         累计器，fDistAccOut 实时镜像，行为一致（镜像同源）；
 *                         ④ 组态闸：润滑里程 <= 0 / 锁定窗 < 0 → 故障锁存；
 *                         ⑤ bLubeReq 置位期间累计器冻结（同窗不重复触发，
 *                         PT 保持时长语义，R219 口径）。
 * 码位     (Codes)      : 按 R297 范式零 16# 码位硬编码；错误出口 BOOL+ENUM(eCause)，
 *                         码位待主控收口统一派号。
 * 红线自检 (Redline)    : 7 项红线已自检：R1 零全局 ✓｜R2 零物理地址 ✓｜R3 纯 IEC ✓
 *                         R4 跳变闸/NaN 拒收/组态闸 ✓｜R5 双语同行注释 ✓
 *                         R6 N/A（监视型无状态机，判据纯派生）✓
 *                         R7 TON/R_TRIG 段 0 无条件刷新 ✓
 * 验收向量 (Acceptance) : V1 fLubeDistMm=1000，位置 0→500→1000 → 第二拍后
 *                         bLubeReq=TRUE，fDistAccOut≈1000；
 *                         V2 位置单拍跳变 5000（限 1000）→ 拒收，nJumpCnt=1；
 *                         V3 bLubeDone 沿 → 里程清零重开窗，锁定窗内不重触发。
 * 修订历史 (Revision)   : 2026-11-20  v1.0.0  R49 首版（批 4 · 序号 19）
 *==============================================================================*)
TYPE E_DL_AltCause :
(
    eNone       := 0,                        (* 无故障成因 / No cause *)
    eCfgIllegal := 1                        (* 组态非法：里程/锁定窗越域 / Illegal config *)
);
END_TYPE

FUNCTION_BLOCK FB_DL_AxisLubeDistTrig
VAR_INPUT
    fPosNow     : LREAL := 0.0;              (* 轴当前位置快照 [mm] / Axis position snapshot *)
    fLubeDistMm : LREAL := 10000.0;          (* 润滑里程窗，域 > 0.0 [mm] / Lube distance window *)
    fJumpLimitMm: LREAL := 100.0;            (* 单拍位置增量上限（跳变判据），域 > 0.0 [mm] / Per-scan jump limit *)
    tLubeLockout: TIME := T#5S;              (* 润滑后最小间隔窗，域 >= T#0S [ms] / Post-lube lockout window *)
    bLubeDone   : BOOL := FALSE;             (* 润滑完成确认，上升沿清里程重开窗 [-] / Lube-done ack edge *)
    bEnable     : BOOL := TRUE;              (* 计程使能，FALSE 冻结累计 [-] / Enable *)
    bReset      : BOOL := FALSE;              (* 复位命令，上升沿清里程/台账/故障 [-] / Reset command *)
END_VAR
VAR_OUTPUT
    bLubeReq    : BOOL;                      (* 润滑请求电平（bLubeDone 沿或复位沿清）[-] / Lube request level *)
    fDistAccOut : LREAL;                     (* 当前窗内累计里程（实时镜像）[mm] / Accumulated distance mirror *)
    fTotalDist  : LREAL;                     (* 总里程累计（维护台账）[mm] / Total distance ledger *)
    nJumpCnt    : UDINT;                     (* 位置跳变拒收累计（信息级台账）[次] / Jump rejection counter *)
    eCause      : E_DL_AltCause;             (* 成因出口（R190 归因唯一） / Cause outlet *)
    bError      : BOOL;                      (* 组态故障锁存标志 [-] / Config fault flag *)
END_VAR
VAR
    rtDone   : R_TRIG;                       (* 润滑完成沿实例，段 0 无条件调用 / Done edge instance *)
    rtReset  : R_TRIG;                       (* 复位沿实例，段 0 无条件调用 / Reset edge instance *)
    tonLock  : TON;                          (* 润滑后锁定窗计时，自复位式 IN := NOT Q（R188） / Lockout timer, self-resetting *)
    _fPosPrev: LREAL;                        (* 上拍位置（增量基准）[mm] / Previous position *)
    _fAcc    : LREAL;                        (* 窗内里程累计器（锁存量，判据源）[mm] / Window distance accumulator *)
    _fTotal  : LREAL;                        (* 总里程累计器（锁存量）[mm] / Total accumulator *)
    _bReq    : BOOL;                         (* 润滑请求锁存位 / Lube request latch *)
    _bLock   : BOOL;                         (* 润滑后锁定门控（锁定窗内禁止再触发）[-] / Post-lube lock gate *)
    _dPos    : LREAL;                        (* 本拍位置增量 [mm] / Position delta this scan *)
    _bFault  : BOOL;                         (* 组态故障锁存位 / Config fault latch bit *)
END_VAR
VAR CONSTANT
    DL_ALT_EPS : LREAL := 1.0E-9;            (* 判零容差（增量/里程比较）[mm] / Zero epsilon *)
END_VAR

(* —— 段 0：沿实例无条件刷新（R228A） —— *)
rtDone(CLK := bLubeDone);                    (* 完成沿每拍必调 / Done edge every scan *)
rtReset(CLK := bReset);                      (* 复位沿每拍必调 / Reset edge every scan *)
tonLock(IN := _bLock, PT := tLubeLockout);   (* 锁定窗计时：IN 由锁定门控派生，段 0 无条件刷新（R228A） / Lockout timer, phase-derived IN *)
IF tonLock.Q THEN
    _bLock := FALSE;                         (* 锁定窗到时：解除门控（每拍全路径派生，R285） / Lockout elapsed: release gate *)
END_IF
_dPos := fPosNow - _fPosPrev;                (* 本拍位置增量派生 / Delta derive *)
_fPosPrev := fPosNow;                        (* 增量基准推进 / Base advance *)
_fPosPrev := fPosNow;                        (* 增量基准推进 / Base advance *)

(* —— 段 1：复位沿处理（作用域：清故障 + 清累计器 ×2 + 清请求锁存 + 清台账 + 基准重锚，R283 逐项声明） —— *)
IF rtReset.Q THEN
    _bFault := FALSE;                        (* 清故障锁存 / Clear fault *)
    eCause := E_DL_AltCause.eNone;           (* 清成因 / Clear cause *)
    _fAcc := 0.0;                            (* 清窗内里程 / Clear window distance *)
    _fTotal := 0.0;                          (* 清总里程 / Clear total *)
    _bReq := FALSE;                          (* 清请求锁存 / Clear request latch *)
    _bLock := FALSE;                         (* 清锁定门控 / Clear lock gate *)
    nJumpCnt := 0;                           (* 清跳变台账 / Clear jump counter *)
    _fPosPrev := fPosNow;                    (* 增量基准重锚（防复位巨增量） / Re-anchor base *)
    bLubeReq := FALSE;                       (* 清请求出口 / Clear request outlet *)
END_IF

(* —— 段 2：组态闸故障锁存（R45 配对；锁存至复位沿，R189） —— *)
IF ((fLubeDistMm <= DL_ALT_EPS) OR (fJumpLimitMm <= DL_ALT_EPS) OR (tLubeLockout < T#0S)
    OR (fLubeDistMm <> fLubeDistMm) OR (fJumpLimitMm <> fJumpLimitMm)) AND NOT _bFault THEN
    _bFault := TRUE;                         (* 组态非法/NaN 锁存 / Latch config fault *)
    eCause := E_DL_AltCause.eCfgIllegal;     (* 成因：组态非法 / Cause: illegal config *)
END_IF

(* —— 段 3：计程与触发（监视型纯派生，无 CASE 相） —— *)
IF bEnable AND NOT _bFault THEN
    IF (fPosNow <> fPosNow) OR ((fPosNow - fPosNow) <> (fPosNow - fPosNow)) THEN
        (* 位置 NaN：增量拒收不累计（边界②），基准已推进防坏值滞留 / NaN: skip *)
        ;                                    (* 空语句：ST 语法要求分支非空，无副作用 / Empty statement, ST syntax requires non-empty branch *)
    ELSIF NOT _bReq THEN                     (* 请求挂起期间累计器冻结（边界⑤同窗不重复触发） / Accumulator frozen while requested *)
        IF ABS(_dPos) > fJumpLimitMm THEN
            nJumpCnt := nJumpCnt + 1;        (* 跳变拒收台账（信息级，不置故障级，R90 口径） / Jump counter, info level *)
        ELSIF ABS(_dPos) > DL_ALT_EPS THEN
            _fAcc := _fAcc + ABS(_dPos);     (* 有效增量入窗累计 / Valid delta accumulate *)
            _fTotal := _fTotal + ABS(_dPos); (* 总里程累计 / Total accumulate *)
            IF _fAcc >= fLubeDistMm THEN
                _bReq := TRUE;               (* 里程到窗：请求锁存至完成沿 / Request latch *)
            END_IF
        END_IF
    END_IF
    IF rtDone.Q AND _bReq THEN               (* 完成沿：清里程重开窗 + 启动锁定门控 / Done edge: clear window, arm lock *)
        _bReq := FALSE;                      (* 清请求锁存 / Clear request *)
        _fAcc := 0.0;                        (* 清窗内里程 / Clear window *)
        _bLock := TRUE;                      (* 锁定门控置位（锁定窗计时由段 0 无条件推进） / Arm lock gate *)
    END_IF
END_IF

(* —— 段 4：出口映射（判据读锁存、镜像同源，红线要求一致行为） —— *)
bLubeReq := _bReq AND NOT _bLock AND (NOT _bFault) AND bEnable;   (* 请求出口：锁存 ∧ 锁定门外 ∧ 非故障 ∧ 使能（锁定窗内收敛防连环请求） / Request outlet with lock gating *)
fDistAccOut := _fAcc;                        (* 窗内里程实时镜像 / Window mirror *)
fTotalDist := _fTotal;                       (* 总里程镜像 / Total mirror *)
bError := _bFault;                           (* 组态故障镜像 / Config fault mirror *)
END_FUNCTION_BLOCK
